(* IEC 61131-3 sources: daoli-st-library/DL_Base (part 2) *)

(* ---- FC_DL_DewPointSurfaceRiskCalc.st ---- *)
(*
  Component : FC_DL_DewPointSurfaceRiskCalc
  Category  : DL_Base
  Function  : 表面结露风险：按 Magnus 公式求露点，与表面温度比较并给出裕度与风险等级
  Complexity: C2
  开源溯源 : DLF 内部原创（R94 族模板派生）；参考语义来源见 SOURCE_HUNTING_MATRIX.md
  规则遵从 : R1-R16
  契约     : 输入 rAmbientC 环境温度 [℃]、rRelHumPct 相对湿度 [%]、rSurfaceC 表面温度 [℃]、
             rMarginWarnK 预警裕度 [K]、rMarginSafeK 安全裕度 [K]；
             输出 rDewPointC 露点温度 [℃]、rMarginK 表面温度减露点 [K]、eRisk 风险等级、
             xValid 有效标志、nFaultCode 故障码。
  边界     : Magnus 系数 a=17.62、b=243.12 [℃]；γ = ln(RH/100) + a·T/(b+T)，露点 Td = b·γ/(a−γ)；
             (a−γ) 为分母须 >1.0E-6（γ 逼近 a 时露点发散）；相对湿度须在 (0,100] [%] 内；
             裕度判级：裕度 < 0 → eRisky（已结露）；< 预警裕度 → eCaution；≥ 安全裕度 → eSafe；
             预警裕度须 ≤ 安全裕度（否则分级区间为空，判 9803）。
  码位     : 9801 输入非有限（故障级）；9802 湿度或分母越域（故障级）；9803 裕度配比越域（故障级）。
*)
TYPE E_DL_DewRisk :
(
    eSafe    := 0,    // 安全：裕度不小于安全裕度 EN: safe, the margin reaches the safe margin
    eCaution := 1,    // 预警：裕度在预警与安全之间 EN: caution, the margin sits between the two limits
    eRisky   := 2     // 危险：裕度不足或已结露 EN: risky, the margin is insufficient or condensation already occurs
);
END_TYPE

FUNCTION FC_DL_DewPointSurfaceRiskCalc : BOOL
VAR_INPUT
    rAmbientC    : LREAL := 30.0;    // 环境温度 [℃] EN: the ambient temperature
    rRelHumPct   : LREAL := 60.0;    // 相对湿度 [%] EN: the relative humidity
    rSurfaceC    : LREAL := 25.0;    // 表面温度 [℃] EN: the surface temperature
    rMarginWarnK : LREAL := 2.0;     // 预警裕度 [K] EN: the warning margin
    rMarginSafeK : LREAL := 5.0;     // 安全裕度 [K] EN: the safe margin
END_VAR
VAR_OUTPUT
    rDewPointC : LREAL;              // 露点温度 [℃] EN: the dew point temperature
    rMarginK   : LREAL;              // 表面温度减露点 [K] EN: the surface temperature minus the dew point
    eRisk      : E_DL_DewRisk;       // 风险等级 EN: the condensation risk level
    xValid     : BOOL;               // 输出可信标志 EN: the outputs are valid
    nFaultCode : INT;                // 0=无故障 9801=输入非有限 9802=湿度或分母越域 9803=裕度配比越域 EN: zero none, 9801 non finite, 9802 humidity or divisor out of range, 9803 margin ordering out of range
END_VAR
VAR
    xFinAll : BOOL;                  // 五输入同时有限 EN: all five inputs are finite
    rRHFrac : LREAL;                 // 相对湿度分数 [-] EN: the relative humidity fraction
    rGamma  : LREAL;                 // Magnus 中间量 γ [-] EN: the Magnus intermediate value
    rDen    : LREAL;                 // 分母 a−γ [-] EN: the divisor, the coefficient minus gamma
    rTd     : LREAL;                 // 露点中间值 [℃] EN: the interim dew point
    rMarg   : LREAL;                 // 裕度中间值 [K] EN: the interim margin
END_VAR
VAR CONSTANT
    DL_DSR_Z      : LREAL := 0.0;     // 浮点零常量 EN: the floating point zero constant
    DL_DSR_HUND   : LREAL := 100.0;   // 百分数换算系数 EN: the percent conversion factor
    DL_DSR_A      : LREAL := 17.62;   // Magnus 系数 a [-] EN: the Magnus coefficient a
    DL_DSR_B      : LREAL := 243.12;  // Magnus 系数 b [℃] EN: the Magnus coefficient b
    DL_DSR_MIN    : LREAL := 1.0E-6;  // 分母下限 EN: the lower bound of the divisor
    DL_DSR_C_BAD  : INT := 9801;      // 输入非有限 EN: a non finite input
    DL_DSR_C_HUM  : INT := 9802;      // 湿度或分母越域 EN: the humidity or the divisor is out of range
    DL_DSR_C_MARG : INT := 9803;      // 裕度配比越域 EN: the margin ordering is out of range
END_VAR

// 段1｜出口预置
FC_DL_DewPointSurfaceRiskCalc := FALSE;   // 返回值预置假 EN: preset the return value to false
rDewPointC := DL_DSR_Z;                   // 露点预置零 [℃] EN: preset the dew point to zero
rMarginK := DL_DSR_Z;                     // 裕度预置零 [K] EN: preset the margin to zero
eRisk := E_DL_DewRisk.eRisky;             // 风险等级预置为危险（安全侧缺省） EN: preset the risk to risky on the safe side
xValid := FALSE;                          // 有效标志预置假 EN: preset the validity flag to false
nFaultCode := 0;                          // 故障码预置零 EN: preset the fault code to zero

// 段2｜非有限闸：五输入全列
xFinAll := (rAmbientC = rAmbientC) AND ((rAmbientC - rAmbientC) = DL_DSR_Z)
        AND (rRelHumPct = rRelHumPct) AND ((rRelHumPct - rRelHumPct) = DL_DSR_Z)
        AND (rSurfaceC = rSurfaceC) AND ((rSurfaceC - rSurfaceC) = DL_DSR_Z)
        AND (rMarginWarnK = rMarginWarnK) AND ((rMarginWarnK - rMarginWarnK) = DL_DSR_Z)
        AND (rMarginSafeK = rMarginSafeK) AND ((rMarginSafeK - rMarginSafeK) = DL_DSR_Z);   // 五输入有限性 EN: the finiteness of all five inputs
IF NOT xFinAll THEN                                                                          // 非有限出口 EN: leave early on a non finite input
    nFaultCode := DL_DSR_C_BAD;                                                              // 非有限码 EN: the non finite code
    RETURN;                                                                                  // 早退 EN: return early
END_IF

// 段3｜域闸：湿度 (0,100]、裕度配比 预警 ≤ 安全、Magnus 分母 b+T 必须远离零点
IF (rRelHumPct <= DL_DSR_Z) OR (rRelHumPct > DL_DSR_HUND) THEN                                // 湿度域闸 EN: the humidity domain gate
    nFaultCode := DL_DSR_C_HUM;                                                              // 湿度越域码 EN: the humidity code
    RETURN;                                                                                  // 早退 EN: return early
END_IF
IF (DL_DSR_B + rAmbientC) < DL_DSR_MIN THEN                                                   // b+T 分母闸（防 −243.12 ℃ 处除零） EN: guard the b plus T divisor
    nFaultCode := DL_DSR_C_HUM;                                                              // 越域码 EN: the out of range code
    RETURN;                                                                                  // 早退 EN: return early
END_IF
IF (rMarginWarnK > rMarginSafeK) OR (rMarginWarnK < DL_DSR_Z) THEN                            // 裕度配比闸 EN: the margin ordering gate
    nFaultCode := DL_DSR_C_MARG;                                                             // 配比越域码 EN: the margin ordering code
    RETURN;                                                                                  // 早退 EN: return early
END_IF

// 段4｜主体：Magnus 露点
rRHFrac := rRelHumPct / DL_DSR_HUND;                                                          // 湿度分数 [-] EN: the humidity fraction
rGamma := LN(rRHFrac) + (DL_DSR_A * rAmbientC) / (DL_DSR_B + rAmbientC);                      // γ [-]，分母 b+T 在工程域内恒正 EN: the Magnus intermediate
rDen := DL_DSR_A - rGamma;                                                                    // 分母 a−γ [-] EN: the divisor
IF ABS(rDen) < DL_DSR_MIN THEN                                                                // 分母下限保护 EN: guard the divisor
    nFaultCode := DL_DSR_C_HUM;                                                               // 越域码 EN: the out of range code
    RETURN;                                                                                   // 早退 EN: return early
END_IF
rTd := (DL_DSR_B * rGamma) / rDen;                                                            // 露点 [℃] EN: the dew point
IF rTd <> rTd THEN                                                                            // 结果复检 EN: recheck the result
    nFaultCode := DL_DSR_C_HUM;                                                               // 复检失败码 EN: the recheck failure code
    RETURN;                                                                                   // 早退，出口保持零哨兵 EN: return early with the zero sentinels
END_IF

// 段5｜裕度与分级：先算裕度再分级（分级只依赖裕度与两个限值，单源赋值）
// 两个限值已在段3 完成域闸，故分级区间不会出现空集 EN: the two limits passed the gate in section three, so the bands are never empty
rMarg := rSurfaceC - rTd;                                                                     // 裕度 [K] EN: the margin
IF rMarg < DL_DSR_Z THEN                                                                      // 已结露 EN: condensation already occurs
    eRisk := E_DL_DewRisk.eRisky;                                                             // 危险 EN: risky
ELSIF rMarg < rMarginWarnK THEN                                                               // 低于预警裕度 EN: below the warning margin
    eRisk := E_DL_DewRisk.eRisky;                                                             // 危险 EN: risky
ELSIF rMarg < rMarginSafeK THEN                                                               // 预警区间 EN: the caution band
    eRisk := E_DL_DewRisk.eCaution;                                                           // 预警 EN: caution
ELSE
    eRisk := E_DL_DewRisk.eSafe;                                                              // 安全 EN: safe
END_IF

// 段6｜出口
rDewPointC := rTd;                                                                            // 露点出口 [℃] EN: the dew point output
rMarginK := rMarg;                                                                            // 裕度出口 [K] EN: the margin output
xValid := TRUE;                                                                               // 结果可信 EN: the results are valid
FC_DL_DewPointSurfaceRiskCalc := TRUE;                                                        // 返回真 EN: return true
END_FUNCTION

(* ---- FC_DL_DwRealReinterp.st ---- *)
// FC_DL_DwRealReinterp v1.0.0
// 开源溯源：brOscatLib / URL https://github.com/iec-oscat-mirror / 许可证 MIT / 借鉴 DW_TO_REAL+REAL_TO_DW 位重解释语义（双向往返单件），clean-room 重写
(*
  道莅工业代码库 | DL_Base | FC_DL_DwRealReinterp
  版本: 1.0.0 | 日期: 2026-11-23 | 轮次: R75
  功能: DWORD↔REAL IEEE-754 单精度位重解释，双向单件（eMode 选择方向）。
        不用 UNION/POINTER/AT，纯标准移位/掩码手工打包解包（R3 红线口径）
  邻件关系: 全库无位重解释属主（查重留痕 §3 驳回 9 条注）；与 SwapBytes16/32
            字节序族互不重叠（字节序 vs 位级重解释）
  精度边界: 打包方向次正规数钳位为零（bClamped 置位）；Inf/NaN 拒收置码；
            解包方向 e=0 次正规/零按 0 返回，e=255 Inf/NaN 拒收置码
*)
TYPE E_DL_DwRealDir :
(
    eRealToDw := 0,   // REAL → DWORD 打包 / Pack REAL to DWORD bits
    eDwToReal := 1    // DWORD → REAL 解包 / Unpack DWORD bits to REAL
);
END_TYPE

FUNCTION FC_DL_DwRealReinterp : REAL
VAR_INPUT
    fValue : REAL  := 0.0;                        // REAL 方向输入值（eMode=打包时用）/ REAL input for pack direction
    dwBits : DWORD := 16#0000_0000;               // DWORD 方向输入位型（eMode=解包时用）/ DWORD input for unpack direction
    eMode  : E_DL_DwRealDir := E_DL_DwRealDir.eRealToDw;   // 方向选择 / Direction selector
END_VAR
VAR_OUTPUT
    dwOut     : DWORD;                            // 打包输出位型 / Packed DWORD output
    fOut      : REAL;                             // 解包输出值 / Unpacked REAL output
    bValid    : BOOL;                             // 结果有效回执 [-] / Result validity receipt
    bClamped  : BOOL;                             // 次正规数钳位标志 [-] / Subnormal clamped flag
    uErrorId  : UDINT;                            // 事件码，0 = 无事件；16#0002_1B01 = 非有限拒收 / Event code
END_VAR
VAR CONSTANT
    DL_DWR_MANT_SHL : DWORD := 16#007F_FFFF;      // 尾数掩码（低 23 位）/ Mantissa mask, low 23 bits
    DL_DWR_EXP_SHL  : DWORD := 16#7F80_0000;      // 指数掩码（位 30..23）/ Exponent mask, bits 30..23
    DL_DWR_SIGN_SHL : DWORD := 16#8000_0000;      // 符号位掩码 / Sign bit mask
    DL_DWR_EXPONE   : DWORD := 16#3F80_0000;      // 指数=127（1.0 尾数基位）/ Exponent 127, mantissa 1.0 base
    DL_DWR_ABSMIN   : REAL := 1.18E-38;           // 最小正规数阈值 [无量纲] / Min normal magnitude
    DL_DWR_ABSMAX   : REAL := 3.40E38;            // 最大可表幅值阈值 [无量纲] / Max representable magnitude
END_VAR
VAR
    fAbs   : REAL;                                // 输入幅值 [无量纲] / Input magnitude
    bNeg   : BOOL;                                // 符号位 [-] / Sign flag
    fExpF  : REAL;                                // 实数域指数中间量 [1] / Real-domain exponent intermediate
    nExp   : INT;                                 // 偏置指数（域 0..254）[1] / Biased exponent, 0..254
    fMant  : REAL;                                // 尾数份额 ∈ [0,1) [1] / Mantissa fraction in [0,1)
    dwMant : DWORD;                               // 尾数位型（23 位）/ Mantissa bits
    dwExp  : DWORD;                               // 指数位型 / Exponent bits
    dwSign : DWORD;                               // 符号位型 / Sign bits
    dwAll  : DWORD;                               // 组合位型 / Combined bits
    nExpU  : INT;                                 // 解包方向指数 [1] / Unpack exponent
    fTwoE  : REAL;                                // 2^nExp 缩放因子 [1] / Scaling factor 2^nExp
    fNorm  : REAL;                                // 归一尾数值 ∈ [1,2) [1] / Normalized mantissa value
    i      : INT;                                 // 指数迭代计数 [次] / Exponent iteration counter
    dwM    : DWORD;                               // 解包方向尾数位型 / Unpack mantissa bits
    fM     : REAL;                                // 解包方向尾数份额 [1] / Unpack mantissa fraction
END_VAR

// —— 段 0：全路径缺省 —— //
bValid   := FALSE;                              // 有效回执预清 / Validity preset
bClamped := FALSE;                              // 钳位标志预清 / Clamped flag preset
uErrorId := 16#0000;                            // 事件码预清 / Event code preset
dwOut    := 16#0000_0000;                       // 打包输出缺省零位型 / Packed output default
fOut     := 0.0;                                // 解包输出缺省零 / Unpacked output default
FC_DL_DwRealReinterp := 0.0;                    // 返回值缺省零（解包方向结果镜像）/ Return default mirrors unpack result

// —— 段 1：方向分派（CASE 全枚举 + ELSE 兜底） —— //
CASE eMode OF

E_DL_DwRealDir.eRealToDw :
    // —— 打包方向：REAL → IEEE-754 位型 —— //
    IF (fValue <> fValue) OR (ABS(fValue) > DL_DWR_ABSMAX) THEN
        uErrorId := 16#0002_1B01;               // 非有限或超可表幅值：拒收置码 / Non-finite or beyond range: reject
        RETURN;
    END_IF
    IF fValue = 0.0 THEN                        // 零（含 -0.0）特判 / Zero special case
        dwOut := 16#0000_0000;                  // 零位型 / Zero bits
        bValid := TRUE;                         // 有效回执 / Validity receipt
        FC_DL_DwRealReinterp := 0.0;            // 返回零 / Return zero
        RETURN;
    END_IF
    fAbs := ABS(fValue);                        // 幅值派生 / Magnitude
    IF fAbs < DL_DWR_ABSMIN THEN                // 次正规域：钳位为零（本件精度边界）/ Subnormal domain: clamp to zero
        bClamped := TRUE;                       // 钳位标志 / Clamped flag
        dwOut := 16#0000_0000;                  // 零位型 / Zero bits
        bValid := TRUE;                         // 有效（确定行为，不发散）/ Valid, deterministic
        RETURN;
    END_IF
    bNeg := (fValue < 0.0);                     // 符号提取 / Sign extraction
    fExpF := LOG(fAbs) / 0.693147180559945;     // log2(|f|)（ln2 常数除） / log2 of magnitude
    nExp := REAL_TO_DINT(fExpF);                // 截断取整（向零）/ Truncate toward zero
    IF REAL_TO_DINT(fExpF) < 0 THEN             // 负指数截断上偏一格修正 / Negative truncation correction
        IF fExpF < DINT_TO_REAL(nExp) THEN      // 向零截断丢失进位时修正 / Correct when truncation lost carry
            nExp := nExp - 1;                   // 指数下移保证尾数 ∈ [1,2) / Shift exponent so mantissa in [1,2)
        END_IF
    END_IF
    IF nExp < -126 THEN
        nExp := -126;                           // 指数下限钳位 / Exponent lower clamp
    END_IF
    IF nExp > 127 THEN
        nExp := 127;                            // 指数上限钳位 / Exponent upper clamp
    END_IF
    fTwoE := 1.0;                               // 2^nExp 迭代初值 / Iteration base for 2^nExp
    IF nExp >= 0 THEN
        FOR i := 1 TO nExp DO                    // 正指数迭代乘 2 / Positive exponent iteration
            fTwoE := fTwoE * 2.0;
        END_FOR
    ELSE
        FOR i := 1 TO (-nExp) DO                 // 负指数迭代除 2 / Negative exponent iteration
            fTwoE := fTwoE * 0.5;
        END_FOR
    END_IF
    fNorm := fAbs / fTwoE;                      // 归一尾数 ∈ [1,2) / Normalized mantissa
    IF fNorm >= 2.0 THEN                        // LOG 取整舍入上溢一格修正 / Rounding overshoot correction
        fNorm := fNorm * 0.5;                   // 尾数减半，指数加一 / Halve mantissa, bump exponent
        nExp := nExp + 1;
        IF nExp > 127 THEN
            nExp := 127;                        // 指数上限复钳位 / Exponent re-clamp upper
        END_IF
    END_IF
    fMant := fNorm - 1.0;                       // 小数份额 ∈ [0,1) / Fractional part
    dwMant := REAL_TO_DWORD(fMant * 8388608.0); // 份额 ×2^23 取整为位型 / Fraction scaled to 23-bit bits
    dwMant := SHL(dwMant, 0) AND DL_DWR_MANT_SHL;   // 低 23 位掩码（SHL 0 防方言化）/ Mask low 23 bits
    dwExp := DINT_TO_DWORD(nExp + 127);         // 偏置指数位型 / Biased exponent bits
    dwExp := SHL(dwExp, 23) AND DL_DWR_EXP_SHL; // 移位至位 30..23 并掩码 / Shift to bits 30..23 and mask
    IF bNeg THEN
        dwSign := DL_DWR_SIGN_SHL;              // 负号置符号位 / Negative sets sign bit
    ELSE
        dwSign := 16#0000_0000;                 // 正号零位型 / Positive zero bits
    END_IF
    dwOut := dwSign OR dwExp OR dwMant;         // 三段位或组合 / Combine three fields
    bValid := TRUE;                             // 有效回执 / Validity receipt
    FC_DL_DwRealReinterp := 0.0;                // 打包方向返回值无意义，置零 / Return meaningless in pack direction

E_DL_DwRealDir.eDwToReal :
    // —— 解包方向：IEEE-754 位型 → REAL —— //
    IF (dwBits AND DL_DWR_EXP_SHL) = DL_DWR_EXP_SHL THEN     // 指数全 1：Inf/NaN 域 / All-ones exponent: Inf or NaN
        uErrorId := 16#0002_1B01;               // 非有限拒收置码 / Non-finite reject code
        RETURN;
    END_IF
    dwM := dwBits AND DL_DWR_MANT_SHL;          // 尾数位型 / Mantissa bits
    fM := DWORD_TO_REAL(SHR(dwM, 0)) / 8388608.0;   // 尾数份额 ∈ [0,1)（SHR 0 保类型）/ Mantissa fraction
    nExpU := DWORD_TO_DINT(SHR(dwBits AND DL_DWR_EXP_SHL, 23)) - 127;   // 无偏指数 / Unbiased exponent
    IF (nExpU = -127) AND (dwM = 16#0000_0000) THEN          // e=0 且尾数=0：真零 / e=0 with zero mantissa: true zero
        IF (dwBits AND DL_DWR_SIGN_SHL) <> 16#0000_0000 THEN // 负零位型 / Negative zero bits
            fOut := 0.0;                        // 负零按零返回 / Return zero
        ELSE
            fOut := 0.0;                        // 正零 / Positive zero
        END_IF
        bValid := TRUE;                         // 有效回执 / Validity receipt
        FC_DL_DwRealReinterp := fOut;           // 返回镜像 / Return mirror
        RETURN;
    END_IF
    IF nExpU = -127 THEN                        // e=0 且尾数非零：次正规（本件精度边界）/ e=0 nonzero mantissa: subnormal
        bClamped := TRUE;                       // 钳位标志 / Clamped flag
        fOut := 0.0;                            // 次正规按零返回（确定行为）/ Subnormal as zero
        bValid := TRUE;                         // 有效（确定行为）/ Valid
        FC_DL_DwRealReinterp := fOut;           // 返回镜像 / Return mirror
        RETURN;
    END_IF
    fTwoE := 1.0;                               // 2^nExpU 迭代初值 / Iteration base
    IF nExpU >= 0 THEN
        FOR i := 1 TO nExpU DO                   // 正指数迭代 / Positive iteration
            fTwoE := fTwoE * 2.0;
        END_FOR
    ELSE
        FOR i := 1 TO (-nExpU) DO                // 负指数迭代 / Negative iteration
            fTwoE := fTwoE * 0.5;
        END_FOR
    END_IF
    fOut := (1.0 + fM) * fTwoE;                 // (1+mantissa)·2^e / Normalized value
    IF (dwBits AND DL_DWR_SIGN_SHL) <> 16#0000_0000 THEN     // 符号还原 / Sign restore
        fOut := -fOut;                          // 负值 / Negative value
    END_IF
    dwOut := 16#0000_0000;                      // 解包方向打包输出无效，置零位型 / Pack output meaningless here
    bValid := TRUE;                             // 有效回执 / Validity receipt
    FC_DL_DwRealReinterp := fOut;               // 返回值 = 解包结果（调用便利）/ Return equals unpack result

ELSE
    // —— 非法枚举兜底 —— //
    uErrorId := 16#0002_1B01;                   // 信息级：模式非法 / Info level: illegal mode
    RETURN;                                     // 全缺省返回 / Return all defaults
END_CASE
END_FUNCTION

(* ---- FC_DL_EnthalpyUnitConvert.st ---- *)
(*
  FC_DL_EnthalpyUnitConvert —— 比焓换算 kJ/kg 与 kcal/kg 与 BTU/lb
  分类：DL_Base | 复杂度：1 | 轮次：R86
  开源溯源：道莅原创（clean-room 自研，纯 IEC 61131-3 通用算法），无外部代码引用
  许可证：MIT
  职责：把三种比焓单位统一折算到基准单位 kJ/kg（1 kcal/kg = 4.1868 kJ/kg；1 BTU/lb = 2.326 kJ/kg）。
  契约：fIn 输入值 [源单位]，eUnit 源单位枚举；fOut 折算结果 [kJ/kg]；返回 TRUE 表示 fOut 可信。
  边界：未知枚举 / 非有限输入（NaN 自反判、Inf 用 1.0E30 绝对上限判）→ 返回 FALSE，fOut 给 0.0 哨兵；
        无除法（纯乘法定标），零全局、零物理地址、零库件依赖。
*)

(*-----------------------------------------------------------------------------
 * 枚举: E_DL_EnthUnit（比焓单位，归属本文件，全库唯一定义）
 *----------------------------------------------------------------------------*)
TYPE E_DL_EnthUnit :
(
    eKjPerKg   := 0,   // 千焦每千克（基准单位） [kJ/kg] / Kilojoule per kilogram, the base unit
    eKcalPerKg := 1,   // 千卡每千克 [kcal/kg] / Kilocalorie per kilogram
    eBtuPerLb  := 2    // 英热单位每磅 [BTU/lb] / British thermal unit per pound
);
END_TYPE

FUNCTION FC_DL_EnthalpyUnitConvert : BOOL
VAR_INPUT
    fIn   : LREAL := 0.0;              // 输入值 [源单位] / The input value in the source unit
    eUnit : E_DL_EnthUnit;             // 源单位枚举 [—] / The source unit enumeration
END_VAR
VAR_OUTPUT
    fOut : LREAL;                      // 折算结果 [kJ/kg] / The converted value in the base unit
END_VAR
VAR CONSTANT
    DL_EU_KCAL : LREAL := 4.1868;      // 1 kcal/kg 折 kJ/kg 的系数 [-] / kcal per kg to kJ per kg
    DL_EU_BTU  : LREAL := 2.326;       // 1 BTU/lb 折 kJ/kg 的系数 [-] / BTU per lb to kJ per kg
    DL_EU_INF  : LREAL := 1.0E30;      // 非有限 / 越界判据上限 [-] / The magnitude gate
    DL_EU_Z    : LREAL := 0.0;         // 浮点零常量 [kJ/kg] / The floating point zero constant
END_VAR

FC_DL_EnthalpyUnitConvert := FALSE;                       // 返回值预置假 / preset the return false
fOut := DL_EU_Z;                                          // 输出预置零哨兵 [kJ/kg] / preset the zero sentinel
IF (fIn <> fIn) OR (ABS(fIn) > DL_EU_INF) THEN            // 自反判 NaN 或越限判 Inf / NaN or Inf
    fOut := DL_EU_Z;                                      // 非有限值输出零哨兵 [kJ/kg] / zero the non finite input
ELSE
    CASE eUnit OF
        E_DL_EnthUnit.eKjPerKg:                           // 基准单位直通 / the base unit passes through
            fOut := fIn;                                  // 直通不换算 [kJ/kg] / pass through unchanged
            FC_DL_EnthalpyUnitConvert := TRUE;            // 结果可信 / the result is valid
        E_DL_EnthUnit.eKcalPerKg:                         // 千卡每千克 / kilocalorie per kilogram
            fOut := fIn * DL_EU_KCAL;                     // 乘 4.1868 [kJ/kg] / multiply by the factor
            FC_DL_EnthalpyUnitConvert := TRUE;            // 结果可信 / the result is valid
        E_DL_EnthUnit.eBtuPerLb:                          // 英热单位每磅 / British thermal unit per pound
            fOut := fIn * DL_EU_BTU;                      // 乘 2.326 [kJ/kg] / multiply by the factor
            FC_DL_EnthalpyUnitConvert := TRUE;            // 结果可信 / the result is valid
    ELSE
        fOut := DL_EU_Z;                                  // 未知枚举输出零哨兵 [kJ/kg] / zero sentinel on an unknown unit
        FC_DL_EnthalpyUnitConvert := FALSE;               // 未知枚举不可信 / an unknown unit is not valid
    END_CASE
END_IF
END_FUNCTION

(* ---- FC_DL_HeatFluxUnitConvert.st ---- *)
(*
  FC_DL_HeatFluxUnitConvert —— 热流密度换算 W/m2 与 kcal/(h*m2)
  分类：DL_Base | 复杂度：2 | 轮次：R86
  开源溯源：道莅原创（clean-room 自研，纯 IEC 61131-3 通用算法），无外部代码引用
  许可证：MIT
  职责：把热流密度统一折算到基准单位 W/m2（1 kcal/(h*m2) = 1.163 W/m2）。
  契约：fIn 输入值 [源单位]，eUnit 源单位枚举；fOut 折算结果 [W/m2]；返回 TRUE 表示 fOut 可信。
  边界：未知枚举 / 非有限输入 → 返回 FALSE，fOut 给 0.0 哨兵；无除法，零全局、零物理地址、零库件依赖。
*)

(*-----------------------------------------------------------------------------
 * 枚举: E_DL_HfxUnit（热流密度单位，归属本文件，全库唯一定义）
 *----------------------------------------------------------------------------*)
TYPE E_DL_HfxUnit :
(
    eWattPerM2    := 0,   // 瓦每平方米（基准单位） [W/m2] / Watt per square metre, the base unit
    eKcalPerHM2   := 1    // 千卡每小时平方米 [kcal/(h*m2)] / Kilocalorie per hour square metre
);
END_TYPE

FUNCTION FC_DL_HeatFluxUnitConvert : BOOL
VAR_INPUT
    fIn   : LREAL := 0.0;              // 输入值 [源单位] / The input value in the source unit
    eUnit : E_DL_HfxUnit;              // 源单位枚举 [—] / The source unit enumeration
END_VAR
VAR_OUTPUT
    fOut : LREAL;                      // 折算结果 [W/m2] / The converted value in the base unit
END_VAR
VAR CONSTANT
    DL_HF_KCAL : LREAL := 1.163;       // 1 kcal/(h*m2) 折 W/m2 的系数 [-] / kcal per hour square metre to watt per square metre
    DL_HF_INF  : LREAL := 1.0E30;      // 非有限 / 越界判据上限 [-] / The magnitude gate
    DL_HF_Z    : LREAL := 0.0;         // 浮点零常量 [W/m2] / The floating point zero constant
END_VAR

FC_DL_HeatFluxUnitConvert := FALSE;                       // 返回值预置假 / preset the return false
fOut := DL_HF_Z;                                          // 输出预置零哨兵 [W/m2] / preset the zero sentinel
IF (fIn <> fIn) OR (ABS(fIn) > DL_HF_INF) THEN            // 自反判 NaN 或越限判 Inf / NaN or Inf
    fOut := DL_HF_Z;                                      // 非有限值输出零哨兵 [W/m2] / zero the non finite input
ELSE
    CASE eUnit OF
        E_DL_HfxUnit.eWattPerM2:                          // 基准单位直通 / the base unit passes through
            fOut := fIn;                                  // 直通不换算 [W/m2] / pass through unchanged
            FC_DL_HeatFluxUnitConvert := TRUE;            // 结果可信 / the result is valid
        E_DL_HfxUnit.eKcalPerHM2:                         // 千卡每小时平方米 / kcal per hour square metre
            fOut := fIn * DL_HF_KCAL;                     // 乘 1.163 [W/m2] / multiply by the factor
            FC_DL_HeatFluxUnitConvert := TRUE;            // 结果可信 / the result is valid
    ELSE
        fOut := DL_HF_Z;                                  // 未知枚举输出零哨兵 [W/m2] / zero sentinel on an unknown unit
        FC_DL_HeatFluxUnitConvert := FALSE;               // 未知枚举不可信 / an unknown unit is not valid
    END_CASE
END_IF
END_FUNCTION

(* ---- FC_DL_HtcUnitConvert.st ---- *)
(*
  FC_DL_HtcUnitConvert —— 传热系数换算 W/(m2*K) 与 kcal/(h*m2*C) 与 BTU/(h*ft2*F)
  分类：DL_Base | 复杂度：2 | 轮次：R86
  开源溯源：道莅原创（clean-room 自研，纯 IEC 61131-3 通用算法），无外部代码引用
  许可证：MIT
  职责：把传热系数统一折算到基准单位 W/(m2*K)：
        1 kcal/(h*m2*C) = 1.163 W/(m2*K)；1 BTU/(h*ft2*F) = 5.678263 W/(m2*K)。
  契约：fIn 输入值 [源单位]，eUnit 源单位枚举；fOut 折算结果 [W/(m2*K)]；返回 TRUE 表示 fOut 可信。
  边界：未知枚举 / 非有限输入 → 返回 FALSE，fOut 给 0.0 哨兵；无除法，零全局、零物理地址、零库件依赖。
*)

(*-----------------------------------------------------------------------------
 * 枚举: E_DL_HtcUnit（传热系数单位，归属本文件，全库唯一定义）
 *----------------------------------------------------------------------------*)
TYPE E_DL_HtcUnit :
(
    eWattPerM2K    := 0,   // 瓦每平方米开（基准单位） [W/(m2*K)] / Watt per square metre kelvin, the base unit
    eKcalPerHM2C   := 1,   // 千卡每小时平方米摄氏度 [kcal/(h*m2*C)] / Kilocalorie per hour square metre celsius
    eBtuPerHFt2F   := 2    // 英热单位每小时平方英尺华氏度 [BTU/(h*ft2*F)] / BTU per hour square foot fahrenheit
);
END_TYPE

FUNCTION FC_DL_HtcUnitConvert : BOOL
VAR_INPUT
    fIn   : LREAL := 0.0;              // 输入值 [源单位] / The input value in the source unit
    eUnit : E_DL_HtcUnit;              // 源单位枚举 [—] / The source unit enumeration
END_VAR
VAR_OUTPUT
    fOut : LREAL;                      // 折算结果 [W/(m2*K)] / The converted value in the base unit
END_VAR
VAR CONSTANT
    DL_HT_KCAL : LREAL := 1.163;       // kcal/(h*m2*C) 折 W/(m2*K) 的系数 [-] / kcal to watt per square metre kelvin
    DL_HT_BTU  : LREAL := 5.678263;    // BTU/(h*ft2*F) 折 W/(m2*K) 的系数 [-] / BTU to watt per square metre kelvin
    DL_HT_INF  : LREAL := 1.0E30;      // 非有限 / 越界判据上限 [-] / The magnitude gate
    DL_HT_Z    : LREAL := 0.0;         // 浮点零常量 [W/(m2*K)] / The floating point zero constant
END_VAR

FC_DL_HtcUnitConvert := FALSE;                            // 返回值预置假 / preset the return false
fOut := DL_HT_Z;                                          // 输出预置零哨兵 [W/(m2*K)] / preset the zero sentinel
IF (fIn <> fIn) OR (ABS(fIn) > DL_HT_INF) THEN            // 自反判 NaN 或越限判 Inf / NaN or Inf
    fOut := DL_HT_Z;                                      // 非有限值输出零哨兵 [W/(m2*K)] / zero the non finite input
ELSE
    CASE eUnit OF
        E_DL_HtcUnit.eWattPerM2K:                         // 基准单位直通 / the base unit passes through
            fOut := fIn;                                  // 直通不换算 [W/(m2*K)] / pass through unchanged
            FC_DL_HtcUnitConvert := TRUE;                 // 结果可信 / the result is valid
        E_DL_HtcUnit.eKcalPerHM2C:                        // 千卡每小时平方米摄氏度 / kcal per hour square metre celsius
            fOut := fIn * DL_HT_KCAL;                     // 乘 1.163 [W/(m2*K)] / multiply by the factor
            FC_DL_HtcUnitConvert := TRUE;                 // 结果可信 / the result is valid
        E_DL_HtcUnit.eBtuPerHFt2F:                        // 英热单位每小时平方英尺华氏度 / BTU per hour square foot fahrenheit
            fOut := fIn * DL_HT_BTU;                      // 乘 5.678263 [W/(m2*K)] / multiply by the factor
            FC_DL_HtcUnitConvert := TRUE;                 // 结果可信 / the result is valid
    ELSE
        fOut := DL_HT_Z;                                  // 未知枚举输出零哨兵 [W/(m2*K)] / zero sentinel on an unknown unit
        FC_DL_HtcUnitConvert := FALSE;                    // 未知枚举不可信 / an unknown unit is not valid
    END_CASE
END_IF
END_FUNCTION

(* ---- FC_DL_IntervalMembership.st ---- *)
(*==============================================================================
 * 组件名称 (Component)  : FC_DL_IntervalMembership
 * 所属子库 (Sublibrary) : DL_Base
 * 归属目录 (Directory)  : C:\Library\DL_Base
 * 当前版本 (Version)    : 1.0.0
 * 组件分类 (Category)   : 函数（FUNCTION）· 纯函数 · 开闭区间归属判定
 * 兼容性   (Platform)   : CODESYS 3.5 / TwinCAT 3 / 汇川 InoProShop / 施耐德
 *                         Machine Expert；仅用 Standard.library 的 ABS / MIN，
 *                         无厂商扩展，无实例依赖
 * 功能一句话 (Summary)  : 判定一个实数是否落在指定开闭组合的区间内，并给出到
 *                         最近边界的有符号裕量与恰在边界标志。
 * 功能描述 (Function)   : 工艺窗口有大量半开约定，例如温度 60 到 80 左闭右开、
 *                         压力 0.4 到 0.6 左开右闭。本件把「开闭组合」做成独立
 *                         参数，四种组合各走一条判定支路，边界归属不再靠调用方
 *                         记忆，同一产线各工位判定口径由此统一。
 * 与既有件边界 (Boundary): FC_DL_ToleranceWindow 判单点对称公差带；FC_DL_LimitClassify
 *                         做四阈值五档分级；FC_DL_RangeOverlapCheck 判两个区间的关系。
 *                         本件判「单点与一端点开闭组合区间」的归属，与三者正交。
 * 设计要点 (Key notes)  : ① 有限性前置拦截：非数与非有限值直接判不可信，绝不进入
 *                           比较链（非数参与比较恒为假，会静默判成「不在区间」）；
 *                         ② 端点序校验先于一切比较，倒置区间不返回「看似合理」的假；
 *                         ③ 边界容差双向使用：闭侧把贴近值纳入，开侧把贴近值排除，
 *                           同一容差保证「既报超限又报未到」的临界矛盾不再出现；
 *                         ④ 退化区间单列一条判据，只有双闭组合才含单点；
 *                         ⑤ 纯函数：无内部状态，同入参同结果，可重入。
 * 开源溯源 (Origin)     : 来源标签 lgf-comparator。LGF 为免费闭源发布的公开函数库
 *                         手册，本件仅借鉴其比较器组把「区间判断 / 公差窗口 / 限值」
 *                         三分的分类骨架，以及区间带开闭属性的参数域设计；许可证按
 *                         其发布方条款仅作分类参考，本件零代码行、零注释引用，
 *                         属 clean-room 独立实现。容差策略为本库加严项，LGF 无此概念。
 * 码位说明 (Codes)      : 本件独占信息级码段 16#0001_012B 到 16#0001_012C，纯函数
 *                         无锁存面故不占故障级码；与同族 0125 到 012A 相邻不重叠。
 *                         012B 端点倒置 ｜ 012C 非数或非有限值。
 * 依赖说明 (Depends)    : 无 DL_ 内部依赖；仅 Standard.library 的 ABS / MIN。
 * 红线自检 (Redline)    : 零全局变量表依赖 ｜ 零外部变量声明 ｜ 零物理地址
 *                         纯 IEC 61131-3 ｜ 无除法故无除零面 ｜ 全变量双语同行注释
 *                         状态机 N/A（纯函数）｜ 枚举四成员被分支全覆盖并带兜底
 * 修订历史 (Revision)   : 2026-11-15  v1.0.0  首版入库（Round 12 · 区间判定族）
 *============================================================================*)

(*-----------------------------------------------------------------------------
 * 枚举: E_DL_IntervalKind（归属 DL_Base，与 FC_DL_IntervalMembership 同文件）
 * 含义: 区间的端点开闭组合。编号 0 起跳、段间隔 10，便于后续插值而不破坏既有工程。
 *----------------------------------------------------------------------------*)
TYPE E_DL_IntervalKind :
(
    eClosedClosed := 0,      // 双闭：两端点都计入，退化区间仅此组合包含单点 / Both ends included, only this kind contains a single point
    eClosedOpen   := 10,     // 左闭右开：含下限不含上限，工艺窗口最常见的写法 / Left closed right open, the most common process window
    eOpenClosed   := 20,     // 左开右闭：不含下限含上限 / Left open right closed
    eOpenOpen     := 30      // 双开：两端点都不计入，退化区间为空集 / Both ends excluded, a single point is never inside
);
END_TYPE

(*==============================================================================
 * 判定示意 (Membership picture)：
 *   区间 60 到 80，取值 60 时：左闭组合判在区间内且贴界，左开组合判不在区间内
 *   区间 60 到 80，取值 80 时：右闭组合判在区间内且贴界，右开组合判不在区间内
 *   裕量口径：内正外负，恰在边界为 0；取「到下限距离」与「到上限距离」的较小者
 *   退化区间（上下限相等）：只有双闭组合在贴界时判在区间内，其余三组合恒不在
 *============================================================================*)

(*==============================================================================
 * 逐调用推演 (Call trace)：
 *   调用 1  值 60、下限 60、上限 80、左闭右开
 *     有限性通过；端点有序通过；贴下限为真，贴上限为假
 *     闭侧判据与贴近合取后通过，开侧判据通过，判定在区间内
 *     裕量取 0 与 20 的较小者，得 0，边界标志为真
 *   调用 2  值 80、同区间
 *     贴上限为真；开侧判据为「严格小于且不贴近」，故不通过
 *     判定不在区间内，裕量为 0，边界标志为真（这是本件最重要的语义）
 *   调用 3  值 59.5、同区间
 *     闭侧判据：既不大于等于下限也不贴近，不通过；裕量取 -0.5 与 20.5 的较小者
 *     输出 -0.5，符号自然表达「低于下限」
 *   调用 4  下限 80、上限 60
 *     端点序校验成立（下限大于上限加容差），早退，事件码 012B，判不在区间内
 *============================================================================*)

FUNCTION FC_DL_IntervalMembership : BOOL
VAR_INPUT
    fValue : LREAL;                                             // 被判定值 [工程单位由调用方决定] / Value under test, unit defined by the caller
    fLower : LREAL;                                             // 区间下限 [工程单位由调用方决定] / Lower bound, unit defined by the caller
    fUpper : LREAL;                                             // 区间上限 [工程单位由调用方决定] / Upper bound, unit defined by the caller
    eKind  : E_DL_IntervalKind := E_DL_IntervalKind.eClosedOpen; // 开闭组合，默认左闭右开 / Openness combination, left closed right open by default
    fEps   : LREAL := 1.0E-9;                                   // 边界判定容差，非正时按最小值生效 [工程单位由调用方决定] / Boundary tolerance, non positive falls back to the minimum
END_VAR
VAR_OUTPUT
    bInside     : BOOL;                                         // 落在区间内为真 / Inside the interval
    bOnBoundary : BOOL;                                         // 与某端点距离小于容差为真 / Within tolerance of an endpoint
    fMargin     : LREAL;                                        // 到最近边界的有符号裕量，内正外负，临界为零 [工程单位由调用方决定] / Signed margin to the nearest bound
    uErrorId    : UDINT;                                        // 事件码，0 表示无事件 / Event code, zero means none
    bValid      : BOOL;                                         // 端点有序且三值有限为真 / Bounds ordered and all values finite
END_VAR
VAR
    fEpsUse     : LREAL;                                        // 生效容差，非正输入已回退到最小值 [工程单位由调用方决定] / Effective tolerance after the fallback
    bNearLo     : BOOL;                                         // 贴近下限 / Near the lower bound
    bNearUp     : BOOL;                                         // 贴近上限 / Near the upper bound
    bLoOk       : BOOL;                                         // 下界侧通过 / Lower side passes
    bUpOk       : BOOL;                                         // 上界侧通过 / Upper side passes
    bDegenerate : BOOL;                                         // 退化区间标志，两端点距离小于容差 / Degenerate interval flag
END_VAR
VAR CONSTANT
    DL_EPS_MIN    : LREAL := 1.0E-9;    // 最小容差，容差为零时浮点永不相等故须回退 [工程单位由调用方决定] / Minimum tolerance used when the caller passes zero
    DL_FINITE_MAX : LREAL := 3.4E38;    // 有限性判定上限，超过即视为无穷大 [工程单位由调用方决定] / Finiteness ceiling, beyond this the value counts as infinite
END_VAR

(*------------------------------------------------------------------------------
 * 段 1｜输出预置：任何异常路径下输出确定
 *      Pre-set outputs so that every path is deterministic
 *-----------------------------------------------------------------------------*)
FC_DL_IntervalMembership := FALSE;
bInside                  := FALSE;
bOnBoundary              := FALSE;
fMargin                  := 0.0;
uErrorId                 := 16#0000_0000;
bValid                   := FALSE;

(*------------------------------------------------------------------------------
 * 段 2｜容差归一（边界 B1）：非正容差回退到最小值
 *      Normalise the tolerance: non positive input falls back to the minimum
 *      容差为零时「贴近」判据恒假，闭侧容差与开侧容差同时失效，须显式回退
 *-----------------------------------------------------------------------------*)
fEpsUse := fEps;
IF fEpsUse <= 0.0 THEN
    fEpsUse := DL_EPS_MIN;
END_IF

(*------------------------------------------------------------------------------
 * 段 3｜有限性前置拦截（边界 B2）：非数与无穷大一律判不可信
 *      Non finite interception: NaN and infinity never enter the comparison chain
 *      非数判定用自比较，跨平台一致，不依赖平台扩展函数
 *-----------------------------------------------------------------------------*)
IF (fValue <> fValue) OR (fLower <> fLower) OR (fUpper <> fUpper) THEN
    uErrorId := 16#0001_012C;   // 非数值输入，判定不可信
    RETURN;
END_IF
IF (ABS(fValue) > DL_FINITE_MAX) OR (ABS(fLower) > DL_FINITE_MAX) OR (ABS(fUpper) > DL_FINITE_MAX) THEN
    uErrorId := 16#0001_012C;   // 非有限输入，判定不可信
    RETURN;
END_IF

(*------------------------------------------------------------------------------
 * 段 4｜端点序校验（边界 B3）：倒置区间不返回看似合理的假结果
 *      Endpoint order check: an inverted interval is reported, never guessed
 *-----------------------------------------------------------------------------*)
IF fLower > (fUpper + fEpsUse) THEN
    uErrorId := 16#0001_012B;   // 端点倒置，判不在区间内
    RETURN;
END_IF

(*------------------------------------------------------------------------------
 * 段 5｜边界贴近与退化判定（边界 B4）
 *      Boundary proximity and degeneracy detection
 *-----------------------------------------------------------------------------*)
bNearLo     := ABS(fValue - fLower) < fEpsUse;
bNearUp     := ABS(fValue - fUpper) < fEpsUse;
bOnBoundary := bNearLo OR bNearUp;
bDegenerate := ABS(fUpper - fLower) < fEpsUse;

(*------------------------------------------------------------------------------
 * 段 6｜按开闭组合分派四侧判据（红线：枚举四成员全覆盖并带兜底）
 *      Dispatch the two side checks by the openness combination
 *      闭侧把贴近值纳入，开侧把贴近值排除，同一容差双向使用
 *-----------------------------------------------------------------------------*)
CASE eKind OF

    E_DL_IntervalKind.eClosedClosed:
        bLoOk := (fValue >= fLower) OR bNearLo;
        bUpOk := (fValue <= fUpper) OR bNearUp;

    E_DL_IntervalKind.eClosedOpen:
        bLoOk := (fValue >= fLower) OR bNearLo;
        bUpOk := (fValue < fUpper) AND (NOT bNearUp);

    E_DL_IntervalKind.eOpenClosed:
        bLoOk := (fValue > fLower) AND (NOT bNearLo);
        bUpOk := (fValue <= fUpper) OR bNearUp;

    E_DL_IntervalKind.eOpenOpen:
        bLoOk := (fValue > fLower) AND (NOT bNearLo);
        bUpOk := (fValue < fUpper) AND (NOT bNearUp);

    ELSE
        (* 非法枚举值：不做隐式恢复，判不可信并置兜底码 *)
        (* Illegal enumerator: no implicit recovery, report and stay outside *)
        bLoOk    := FALSE;
        bUpOk    := FALSE;
        uErrorId := 16#0001_012C;
        RETURN;

END_CASE

(*------------------------------------------------------------------------------
 * 段 7｜归属合成（边界 B5）：退化区间只被双闭组合包含
 *      Membership composition: only the doubly closed kind contains a point
 *-----------------------------------------------------------------------------*)
IF bDegenerate THEN
    bInside := (eKind = E_DL_IntervalKind.eClosedClosed) AND bOnBoundary;
ELSE
    bInside := bLoOk AND bUpOk;
END_IF

(*------------------------------------------------------------------------------
 * 段 8｜裕量（边界 B6）：取两侧距离的较小者，外侧自然为负
 *      Margin: the smaller of the two distances, negative outside by nature
 *-----------------------------------------------------------------------------*)
fMargin := MIN(fValue - fLower, fUpper - fValue);

(*------------------------------------------------------------------------------
 * 段 9｜收口：走到此处入参全部合法
 *      Close out: reaching this point means every input is legal
 *-----------------------------------------------------------------------------*)
bValid                   := TRUE;
FC_DL_IntervalMembership := bInside;
END_FUNCTION

(* ---- FC_DL_LevelUnitConvert.st ---- *)
(*
  FC_DL_LevelUnitConvert —— 液位换算 m/mm/%，按罐高换算
  分类：DL_Base | 复杂度：1 | 轮次：R86
  开源溯源：道莅原创（clean-room 自研，纯 IEC 61131-3 通用算法），无外部代码引用
  许可证：MIT
  职责：把液位统一折算到基准单位 m：m 直通、mm 乘 0.001、% 按罐高折算（% × 罐高 / 100）。
  契约：fIn 输入值 [源单位]、eUnit 源单位枚举、fTankHeight 罐内有效高度 [m]；fOut 折算结果 [m]；
        返回 TRUE 表示 fOut 可信。% 通道要求 fTankHeight > 0，否则判不可信（不除零）。
  边界：① 除零防护：仅对 100 常量做除法，罐高为 0 时 % 通道直接判不可信；② 未知枚举 / 非有限输入 → FALSE + 0.0；
        ③ 三个浮点入参逐一做非有限闸；零全局、零物理地址、零库件依赖。
*)

(*-----------------------------------------------------------------------------
 * 枚举: E_DL_LvlUnit（液位单位，归属本文件，全库唯一定义）
 *----------------------------------------------------------------------------*)
TYPE E_DL_LvlUnit :
(
    eMeter    := 0,    // 米（基准单位） [m] / Metre, the base unit
    eMilliMeter := 1,  // 毫米 [mm] / Millimetre
    ePercent  := 2     // 百分比（按罐高折算） [%] / Percent of the tank height
);
END_TYPE

FUNCTION FC_DL_LevelUnitConvert : BOOL
VAR_INPUT
    fIn        : LREAL := 0.0;         // 输入值 [源单位] / The input value in the source unit
    eUnit      : E_DL_LvlUnit;         // 源单位枚举 [—] / The source unit enumeration
    fTankHeight : LREAL := 1.0;        // 罐内有效高度（% 通道必需 > 0） [m] / The effective tank height for percent
END_VAR
VAR_OUTPUT
    fOut : LREAL;                      // 折算结果 [m] / The converted value in the base unit
END_VAR
VAR CONSTANT
    DL_LV_MM   : LREAL := 0.001;       // 1 mm 折 m 的系数 [-] / millimetre to metre
    DL_LV_HUND : LREAL := 100.0;       // 百分比满量程分母 [-] / The percent full scale divisor
    DL_LV_INF  : LREAL := 1.0E30;      // 非有限 / 越界判据上限 [-] / The magnitude gate
    DL_LV_EPS  : LREAL := 1.0E-9;      // 罐高判零容差 [-] / The tank height zero tolerance
    DL_LV_Z    : LREAL := 0.0;         // 浮点零常量 [m] / The floating point zero constant
END_VAR

FC_DL_LevelUnitConvert := FALSE;                          // 返回值预置假 / preset the return false
fOut := DL_LV_Z;                                          // 输出预置零哨兵 [m] / preset the zero sentinel
IF (fIn <> fIn) OR (ABS(fIn) > DL_LV_INF) THEN            // 输入自反判 NaN 或越限判 Inf / the input gate
    fOut := DL_LV_Z;                                      // 非有限值输出零哨兵 [m] / zero the non finite input
ELSIF (fTankHeight <> fTankHeight) OR (ABS(fTankHeight) > DL_LV_INF) THEN // 罐高非有限闸 / the tank height gate
    fOut := DL_LV_Z;                                      // 罐高非法输出零哨兵 [m] / zero sentinel on an invalid height
ELSE
    CASE eUnit OF
        E_DL_LvlUnit.eMeter:                              // 基准单位直通 / the base unit passes through
            fOut := fIn;                                  // 直通不换算 [m] / pass through unchanged
            FC_DL_LevelUnitConvert := TRUE;               // 结果可信 / the result is valid
        E_DL_LvlUnit.eMilliMeter:                         // 毫米折米 / millimetre to metre
            fOut := fIn * DL_LV_MM;                       // 乘 0.001 [m] / multiply by the factor
            FC_DL_LevelUnitConvert := TRUE;               // 结果可信 / the result is valid
        E_DL_LvlUnit.ePercent:                            // 百分比按罐高折算 / percent of the tank height
            IF (fTankHeight > DL_LV_EPS) THEN             // 罐高为正才可折算（除零防护） / a positive height is required
                fOut := (fIn / DL_LV_HUND) * fTankHeight; // 先除常量 100 再乘罐高 [m] / divide then multiply
                FC_DL_LevelUnitConvert := TRUE;           // 结果可信 / the result is valid
            ELSE
                fOut := DL_LV_Z;                          // 罐高为零输出零哨兵 [m] / zero sentinel on a zero height
                FC_DL_LevelUnitConvert := FALSE;          // 不可信 / not valid
            END_IF
    ELSE
        fOut := DL_LV_Z;                                  // 未知枚举输出零哨兵 [m] / zero sentinel on an unknown unit
        FC_DL_LevelUnitConvert := FALSE;                  // 未知枚举不可信 / an unknown unit is not valid
    END_CASE
END_IF
END_FUNCTION

(* ---- FC_DL_MapRangePercent.st ---- *)
(*
  FC_DL_MapRangePercent —— 百分比与工程值互映，枚举方向
  分类：DL_Base | 复杂度：1 | 轮次：R86
  开源溯源：道莅原创（clean-room 自研，纯 IEC 61131-3 通用算法），无外部代码引用
  许可证：MIT
  职责：按 eDir 方向做百分比与工程值互映：
        ePctToEng：fIn 视为百分比 0..100，映射到 [fOutMin, fOutMax]；
        eEngToPct：fIn 视为工程量，映射到百分比 0..100（先钳到量程）。
  契约：fIn 输入值、eDir 方向枚举、fEngMin/fEngMax 工程量程端点；fOut 结果 [目标单位]；返回 TRUE 表示可信。
  边界：① 量程退化校验（容差 DL_MP_EPS）；② 除零防护：分母先过退化闸；③ 浮点入参逐一非有限闸；
        ④ CASE 含 ELSE 兜底拦非法方向；零全局、零物理地址、零库件依赖。
*)

(*-----------------------------------------------------------------------------
 * 枚举: E_DL_MapDir（映射方向，归属本文件，全库唯一定义）
 *----------------------------------------------------------------------------*)
TYPE E_DL_MapDir :
(
    ePctToEng := 0,    // 百分比 → 工程值 [—] / Percent to engineering value
    eEngToPct := 1     // 工程值 → 百分比 [—] / Engineering value to percent
);
END_TYPE

FUNCTION FC_DL_MapRangePercent : BOOL
VAR_INPUT
    fIn     : LREAL := 0.0;            // 输入值 [源单位] / The input value in the source unit
    eDir    : E_DL_MapDir;             // 映射方向枚举 [—] / The mapping direction
    fEngMin : LREAL := 0.0;            // 工程量程下端点 [工程单位] / The engineering range low end
    fEngMax : LREAL := 100.0;          // 工程量程上端点 [工程单位] / The engineering range high end
END_VAR
VAR_OUTPUT
    fOut : LREAL;                      // 结果 [目标单位] / The result in the target unit
END_VAR
VAR
    xBad     : BOOL;                   // 参数非法标志 [—] / The parameter invalid flag
    fInClamp : LREAL;                  // 钳位后的输入 [源单位] / The clamped input value
    fEngSpan : LREAL;                  // 工程量程跨度 [工程单位] / The engineering span
END_VAR
VAR CONSTANT
    DL_MP_EPS   : LREAL := 1.0E-9;     // 浮点比较容差 [-] / The floating point comparison tolerance
    DL_MP_INF   : LREAL := 1.0E30;     // 非有限 / 越界判据上限 [-] / The magnitude gate
    DL_MP_Z     : LREAL := 0.0;        // 浮点零常量 [-] / The floating point zero constant
    DL_MP_HUND  : LREAL := 100.0;      // 百分比满量程 [-] / The percent full scale
END_VAR

FC_DL_MapRangePercent := FALSE;                           // 返回值预置假 / preset the return false
fOut := DL_MP_Z;                                          // 输出预置零哨兵 / preset the zero sentinel
xBad := FALSE;                                            // 非法标志预置假 / preset the invalid flag false
IF (fIn <> fIn) OR (ABS(fIn) > DL_MP_INF) THEN            // 输入非有限闸 / the input gate
    xBad := TRUE;                                         // 置非法标志 / raise the invalid flag
END_IF
IF (fEngMin <> fEngMin) OR (ABS(fEngMin) > DL_MP_INF) THEN // 工程下端非有限闸 / the engineering low end gate
    xBad := TRUE;                                         // 置非法标志 / raise the invalid flag
END_IF
IF (fEngMax <> fEngMax) OR (ABS(fEngMax) > DL_MP_INF) THEN // 工程上端非有限闸 / the engineering high end gate
    xBad := TRUE;                                         // 置非法标志 / raise the invalid flag
END_IF
fEngSpan := fEngMax - fEngMin;                            // 工程量程跨度 [工程单位] / the engineering span
IF ABS(fEngSpan) < DL_MP_EPS THEN                         // 量程退化（除零防护） / the degenerate span
    xBad := TRUE;                                         // 置非法标志 / raise the invalid flag
END_IF
IF NOT xBad THEN                                          // 参数全通过才映射 / map only when all parameters pass
    CASE eDir OF
        E_DL_MapDir.ePctToEng:                            // 百分比转工程值 / percent to engineering value
            fInClamp := fIn;                              // 输入接管 [%] / take the input value
            IF fInClamp < DL_MP_Z THEN                    // 百分比低于零 / below zero percent
                fInClamp := DL_MP_Z;                      // 钳到零 [%] / clamp to zero
            END_IF
            IF fInClamp > DL_MP_HUND THEN                 // 百分比高于一百 / above one hundred percent
                fInClamp := DL_MP_HUND;                   // 钳到一百 [%] / clamp to one hundred
            END_IF
            fOut := fEngMin + (fInClamp / DL_MP_HUND) * fEngSpan; // 线性换算（除常量） [工程单位] / the conversion
            FC_DL_MapRangePercent := TRUE;                // 结果可信 / the result is valid
        E_DL_MapDir.eEngToPct:                            // 工程值转百分比 / engineering value to percent
            fInClamp := fIn;                              // 输入接管 [工程单位] / take the input value
            IF fEngSpan > DL_MP_Z THEN                    // 正常量程方向 / the normal span direction
                IF fInClamp < fEngMin THEN                // 低于下端点 / below the low end
                    fInClamp := fEngMin;                  // 钳到下端点 [工程单位] / clamp to the low end
                END_IF
                IF fInClamp > fEngMax THEN                // 高于上端点 / above the high end
                    fInClamp := fEngMax;                  // 钳到上端点 [工程单位] / clamp to the high end
                END_IF
            ELSE                                          // 反向量程 / the reversed span
                IF fInClamp > fEngMin THEN                // 高于下端（反向即越小越远） / above the low end
                    fInClamp := fEngMin;                  // 钳到下端点 [工程单位] / clamp to the low end
                END_IF
                IF fInClamp < fEngMax THEN                // 低于上端点 / below the high end
                    fInClamp := fEngMax;                  // 钳到上端点 [工程单位] / clamp to the high end
                END_IF
            END_IF
            fOut := ((fInClamp - fEngMin) / fEngSpan) * DL_MP_HUND; // 反向换算（分母已证非零） [%] / the conversion
            FC_DL_MapRangePercent := TRUE;                // 结果可信 / the result is valid
    ELSE
        fOut := DL_MP_Z;                                  // 非法方向输出零哨兵 / zero sentinel on an illegal direction
        FC_DL_MapRangePercent := FALSE;                   // 非法方向不可信 / an illegal direction is not valid
    END_CASE
END_IF
END_FUNCTION

(* ---- FC_DL_SaturateAdd.st ---- *)
(*
  FC_DL_SaturateAdd  —  饱和加减运算 / Saturating add and subtract
  分类 Category : DL_Base
  码位 Code     : 16#01_0_00
  版本 Version  : 1.0.0
  来源 Source   : t2-1-lgf-math — IEC 61131-3 标准语义的道莅防御性实现
  溯源 Origin   : clean-room 实现，通用饱和算术语义，未复制任何源码行
  功能 Function : 1) 以 LINT 宽域中间量计算 nInA ± nInB（Add/Sub 两模式），杜绝 DINT 先加后判的回绕静默翻号；
                  2) 结果先与 [nLimitLo, nLimitHi] 组态区间钳制，再与 DINT 可表达域钳制，输出最终 nOut；
                  3) bClamped 指示本调用发生了钳制（每调用无条件重算，无锁存）。
  边界 Boundary : ① nLimitLo > nLimitHi 判组态错置码，输出 nLimitLo（安全侧下界）且 bClamped := TRUE；
                  ② 结果超出 DINT 可表达域时饱和到对应 DINT 极限并 bClamped := TRUE（DINT ± DINT 在 LINT 内必不溢出，此分支为防御性兜底）；
                  ③ eOp 落入未知值由 CASE ELSE 拦截：置码、输出 0、bClamped := TRUE（不猜运算方向）；
                  ④ 解除式自证：bClamped 为每调用重算量，下一调用结果重新落入区间即自动解除（无 bReset、无锁存）；
                  ⑤ 本件为纯函数：无 VAR 记忆量、无定时器、无边沿实例，可离平台编译。
  依赖 Depends  : 仅 Standard.library（无库调用）；枚举 E_DL_SatOp 随本件发布
  码表 Error codes（本件格 01_0_00，子码步进 +0x100）:
    16#0001_0100 信息级：结果被钳制（bClamped = TRUE，不置故障）
    16#0001_0200 故障级：组态非法 nLimitLo > nLimitHi，输出安全侧下界
    16#0001_0300 故障级：运算模式 eOp 非法（CASE ELSE 兜底）

  修订历史 Revision :
    2026-11-18  v1.0.0  R38 首版
*)

TYPE E_DL_SatOp :
(
    eAdd := 0,   // 加法模式 / Addition mode
    eSub := 1    // 减法模式 / Subtraction mode
);
END_TYPE

FUNCTION FC_DL_SaturateAdd : BOOL
VAR_INPUT
    nInA     : DINT;                 // 操作数 A / Operand A
    nInB     : DINT;                 // 操作数 B / Operand B
    eOp      : E_DL_SatOp;           // 运算模式（Add/Sub）/ Operation mode, Add or Sub
    nLimitHi : DINT;                 // 组态上限 [DINT] / Configured upper limit
    nLimitLo : DINT;                 // 组态下限 [DINT] / Configured lower limit
END_VAR
VAR_OUTPUT
    nOut     : DINT;                 // 钳制后结果 / Saturated result
    bClamped : BOOL;                 // 本调用发生钳制 / Clamped on this call, recomputed per call
    nErrId   : UDINT;                // 事件码，0 = 无事件 / Event code, 0 = none
END_VAR
VAR
    liWork : LINT;                  // 宽域中间量（FC 局部临时量，每调用重算，非记忆量）/ Wide scratch, temp per call
END_VAR
VAR CONSTANT
    DL_DINT_HI : LINT := 2147483647;   // DINT 可表达上界 / Expressible DINT upper bound
    DL_DINT_LO : LINT := -2147483648;  // DINT 可表达下界 / Expressible DINT lower bound
END_VAR

(* —— 段 1：单拍量缺省与组态闸（纯函数，每调用重算） —— *)
nOut     := 0;                        // 输出缺省 0
bClamped := FALSE;                    // 钳制标志每调用重算（无锁存，解除式自证）
nErrId   := 16#0000_0000;             // 事件码缺省无事件

IF nLimitLo > nLimitHi THEN
    nOut     := nLimitLo;             // 组态错：输出安全侧下界（规格强制）
    bClamped := TRUE;                 // 组态错视为钳制
    nErrId   := 16#0001_0200;         // 故障级：组态非法
    FC_DL_SaturateAdd := FALSE;       // 返回值：运算未受理
    RETURN;                            // 组态非法不进入运算
END_IF

(* —— 段 2：LINT 宽域运算（禁先 DINT 相加再判溢出） —— *)
CASE eOp OF

E_DL_SatOp.eAdd:
    liWork := LINT(nInA) + LINT(nInB);   // 宽域加法，DINT±DINT 必不溢出 LINT
    FC_DL_SaturateAdd := TRUE;           // 运算已受理

E_DL_SatOp.eSub:
    liWork := LINT(nInA) - LINT(nInB);   // 宽域减法
    FC_DL_SaturateAdd := TRUE;           // 运算已受理

ELSE
    nOut   := 0;                    // 未知模式：输出 0（不猜方向）
    bClamped := TRUE;               // 视为异常钳制
    nErrId := 16#0001_0300;         // 故障级：运算模式非法
    FC_DL_SaturateAdd := FALSE;     // 运算未受理
    RETURN;

END_CASE

(* —— 段 3：先 DINT 可表达域钳制，再组态区间钳制（顺序不可倒置） —— *)
IF liWork > DL_DINT_HI THEN
    liWork   := DL_DINT_HI;         // 超上界：饱和到 DINT 上限
    bClamped := TRUE;               // 钳制标志
    nErrId   := 16#0001_0100;       // 信息级：结果被钳制
ELSIF liWork < DL_DINT_LO THEN
    liWork   := DL_DINT_LO;         // 超下界：饱和到 DINT 下限
    bClamped := TRUE;
    nErrId   := 16#0001_0100;       // 信息级：结果被钳制
END_IF

IF liWork > LINT(nLimitHi) THEN
    liWork   := LINT(nLimitHi);     // 超组态上限：钳到上限
    bClamped := TRUE;
    nErrId   := 16#0001_0100;       // 信息级：结果被钳制
ELSIF liWork < LINT(nLimitLo) THEN
    liWork   := LINT(nLimitLo);     // 低于组态下限：钳到下限
    bClamped := TRUE;
    nErrId   := 16#0001_0100;       // 信息级：结果被钳制
END_IF

(* —— 段 4：出口单点映射 —— *)
nOut := DINT(liWork);               // 宽域结果回落 DINT（已经两段钳制，必在表达域内）

END_FUNCTION

(* ---- FC_DL_SpecificHeatUnitConvert.st ---- *)
(*
  FC_DL_SpecificHeatUnitConvert —— 比热容换算 kJ/(kg*K) 与 BTU/(lb*F)
  分类：DL_Base | 复杂度：1 | 轮次：R86
  开源溯源：道莅原创（clean-room 自研，纯 IEC 61131-3 通用算法），无外部代码引用
  许可证：MIT
  职责：把比热容统一折算到基准单位 kJ/(kg*K)（1 BTU/(lb*F) = 4.1868 kJ/(kg*K)）。
  契约：fIn 输入值 [源单位]，eUnit 源单位枚举；fOut 折算结果 [kJ/(kg*K)]；返回 TRUE 表示 fOut 可信。
  边界：未知枚举 / 非有限输入 → 返回 FALSE，fOut 给 0.0 哨兵；无除法，零全局、零物理地址、零库件依赖。
*)

(*-----------------------------------------------------------------------------
 * 枚举: E_DL_ShcUnit（比热容单位，归属本文件，全库唯一定义）
 *----------------------------------------------------------------------------*)
TYPE E_DL_ShcUnit :
(
    eKjPerKgK  := 0,   // 千焦每千克开（基准单位） [kJ/(kg*K)] / Kilojoule per kilogram kelvin, the base unit
    eBtuPerLbF := 1    // 英热单位每磅华氏度 [BTU/(lb*F)] / British thermal unit per pound fahrenheit
);
END_TYPE

FUNCTION FC_DL_SpecificHeatUnitConvert : BOOL
VAR_INPUT
    fIn   : LREAL := 0.0;              // 输入值 [源单位] / The input value in the source unit
    eUnit : E_DL_ShcUnit;              // 源单位枚举 [—] / The source unit enumeration
END_VAR
VAR_OUTPUT
    fOut : LREAL;                      // 折算结果 [kJ/(kg*K)] / The converted value in the base unit
END_VAR
VAR CONSTANT
    DL_SC_BTU : LREAL := 4.1868;       // 1 BTU/(lb*F) 折 kJ/(kg*K) 的系数 [-] / BTU per lb F to kJ per kg K
    DL_SC_INF : LREAL := 1.0E30;       // 非有限 / 越界判据上限 [-] / The magnitude gate
    DL_SC_Z   : LREAL := 0.0;          // 浮点零常量 [kJ/(kg*K)] / The floating point zero constant
END_VAR

FC_DL_SpecificHeatUnitConvert := FALSE;                   // 返回值预置假 / preset the return false
fOut := DL_SC_Z;                                          // 输出预置零哨兵 [kJ/(kg*K)] / preset the zero sentinel
IF (fIn <> fIn) OR (ABS(fIn) > DL_SC_INF) THEN            // 自反判 NaN 或越限判 Inf / NaN or Inf
    fOut := DL_SC_Z;                                      // 非有限值输出零哨兵 [kJ/(kg*K)] / zero the non finite input
ELSE
    CASE eUnit OF
        E_DL_ShcUnit.eKjPerKgK:                           // 基准单位直通 / the base unit passes through
            fOut := fIn;                                  // 直通不换算 [kJ/(kg*K)] / pass through unchanged
            FC_DL_SpecificHeatUnitConvert := TRUE;        // 结果可信 / the result is valid
        E_DL_ShcUnit.eBtuPerLbF:                          // 英热单位每磅华氏度 / BTU per pound fahrenheit
            fOut := fIn * DL_SC_BTU;                      // 乘 4.1868 [kJ/(kg*K)] / multiply by the factor
            FC_DL_SpecificHeatUnitConvert := TRUE;        // 结果可信 / the result is valid
    ELSE
        fOut := DL_SC_Z;                                  // 未知枚举输出零哨兵 [kJ/(kg*K)] / zero sentinel on an unknown unit
        FC_DL_SpecificHeatUnitConvert := FALSE;           // 未知枚举不可信 / an unknown unit is not valid
    END_CASE
END_IF
END_FUNCTION

(* ---- FC_DL_StringCompareNatural.st ---- *)
(*==============================================================================
 * 组件名称 (Component)  : FC_DL_StringCompareNatural
 * 所属子库 (Sublibrary) : DL_Base
 * 当前版本 (Version)    : 1.0.0
 * 兼容性   (Platform)   : CODESYS 3.5+ / TwinCAT 3 / 汇川 InoProShop / 施耐德 Machine Expert
 *                         仅依赖 IEC 61131-3 标准字符串九函数（LEN / MID / LEFT / CONCAT / DELETE / FIND），零厂商私有库
 * 功能描述 (Function)   : 自然序比较（Human sort / natural sort）。规则：
 *                           · 双方同位置均为数字时，各自提取完整数字段，按「数值」比较
 *                             （去前导零后先比位数、同位数再逐位比较），故 A2 < A10；
 *                           · 其余位置按单字符序数比较，序数由排序字符集常量
 *                             DL_SCN_ORDER 的 FIND 位置给出（集合外字符序数记 0，排最前）；
 *                           · 公共前缀耗尽后，剩余字符多者更大（A < AB）。
 *                         全程用 FIND(集合, 单字符) 取序数，不依赖平台字符串比较运算符或
 *                         字符码强转方言（R3 纯标准函数路径）。
 * 接口     (Interface)  : 输入 sInA 左串、sInB 右串 [-]；
 *                         输出 iResult 比较结果（-1 左小 / 0 相等 / 1 左大）[-]、
 *                         bEqual 是否相等、eErrCode 错误码（E_DL_StrNatErr）；
 *                         返回值 = bValid 比较可信标志（TRUE = iResult 可信）。
 * 边界     (Boundary)   : ① 属主边界：只做比较，不做排序（排序归调用方的数组管理）、
 *                         不做大小写折叠（'A' 与 'a' 序数不同，A 在前）。
 *                         ② 数字段归一：去前导零后 '007' 与 '7' 相等（数值 7），
 *                         故 "A007" = "A7"（iResult=0）；长度差由去零后的位数决定。
 *                         ③ 序数集合只含 0-9 / A-Z / a-z；标点与空格序数记 0（同序则继续后移，
 *                         不判等、不报错），排序稳定性由调用方的稳定排序保证。
 *                         ④ 长度均钳位至 255（缓冲可表性），双向扫描严格有界。
 *                         ⑤ 内层数字段提取循环亦以上界 _udLenA/_udLenB 收口，无越界。
 *                         ⑥ 零全局耦合（无 GVL / VAR_EXTERNAL / 物理地址）。
 * 分工声明 (Scope)      : 与 `FC_DL_StringReverse` 分工：位序重排归那件、序比较归本件；
 *                         与 `FC_DL_StringIsNumeric` 分工：整串数值判定归那件。
 * 来源标签 (Source Tag) : 原创实现（无外部代码引入）
 * 码表     (Codes)      : 本件不占用全局数字码位；出口为 BOOL + INT + BOOL +
 *                         本文件内定义 enum E_DL_StrNatErr（全库唯一）。
 * 红线自检 (Redline)    : R1 ✓ 零 GVL/VAR_EXTERNAL ｜ R2 ✓ 零 %I/%Q/%M ｜ R3 ✓ 纯 IEC 61131-3
 *                         R4 ✓ 双层循环上界收口 + 去前导零守恒 + 序数集合法（无字符码强转） ｜ R5 ✓ 声明逐行同行双语注释
 *                         R6 N/A（纯函数无状态机） ｜ R7 N/A（无实例调用）
 * 修订历史 (Revision)   : 2026-11-23  v1.0.0  R77 首版（批次 B2 · 序号 9）
 * 验收向量 (Acceptance) : ① sInA='A2', sInB='A10' → iResult=-1（数字段 2 < 10）, bEqual=FALSE, eOk；
 *                         ② sInA='A2', sInB='A2' → iResult=0, bEqual=TRUE；
 *                         ③ sInA='A007', sInB='A7' → 去零后数值相同 → iResult=0, bEqual=TRUE；
 *                         ④ sInA='A', sInB='AB' → 公共前缀耗尽，右串剩余 → iResult=-1；
 *                         ⑤ sInA='B1', sInB='A99' → 首字符序数 B > A → iResult=1；
 *                         ⑥ sInA='', sInB='' → iResult=0, bEqual=TRUE, eOk。
 *==============================================================================*)

(*-----------------------------------------------------------------------------
 * 枚举: E_DL_StrNatErr（自然序比较错误码，归属 DL_Base，与本件同文件，全库唯一属主）
 *----------------------------------------------------------------------------*)
TYPE E_DL_StrNatErr :
(
    eOk      := 0,   // 信息级：比较完成，结果可信 / Info: comparison completed, result trustworthy
    eClampLen:= 1    // 信息级：输入超缓冲上限已按 255 字符比较 / Info: inputs clamped to 255 chars for comparison
);
END_TYPE

FUNCTION FC_DL_StringCompareNatural : BOOL
VAR_INPUT
    sInA : STRING(255);   // 左串 [-] / Left string
    sInB : STRING(255);   // 右串 [-] / Right string
END_VAR
VAR_OUTPUT
    iResult : INT;        // 比较结果：-1 左小 / 0 相等 / 1 左大 [-] / Compare result: -1 less, 0 equal, 1 greater
    bEqual  : BOOL;       // 是否相等（iResult=0） [-] / Whether equal, iResult equals zero
    eErrCode: E_DL_StrNatErr; // 错误码出口 [-] / Error code outlet
END_VAR
VAR
    _udLenA  : UDINT;       // 左串生效长度 [字符] / Effective left length [chars]
    _udLenB  : UDINT;       // 右串生效长度 [字符] / Effective right length [chars]
    _udA     : UDINT;       // 左串游标（1 基） [-] / Left cursor, 1-based
    _udB     : UDINT;       // 右串游标（1 基） [-] / Right cursor, 1-based
    _udKa    : UDINT;       // 数字段内位序 [-] / Bit index inside digit run
    _udRunA  : UDINT;       // 左数字段长度 [字符] / Left digit run length [chars]
    _udRunB  : UDINT;       // 右数字段长度 [字符] / Right digit run length [chars]
    _rkA     : UDINT;       // 左字符序数（0 = 集合外） [-] / Left character rank, 0 means outside set
    _rkB     : UDINT;       // 右字符序数（0 = 集合外） [-] / Right character rank, 0 means outside set
    _sChA    : STRING(255); // 左串当前单字符 [-] / Current left character
    _sChB    : STRING(255); // 右串当前单字符 [-] / Current right character
    _sRunA   : STRING(255); // 左数字段（已去前导零） [-] / Left digit run, leading zeros stripped
    _sRunB   : STRING(255); // 右数字段（已去前导零） [-] / Right digit run, leading zeros stripped
    _iRes    : INT;         // 比较结果内部累加 [-] / Internal compare result
END_VAR
VAR CONSTANT
    DL_SCN_SET_DIGIT : STRING(255) := '0123456789';   // 数字字符集 [-] / Digit character set
    DL_SCN_SET_ZERO  : STRING(255) := '0';            // 零字符集（去前导零用） [-] / Zero character set for leading-zero strip
    DL_SCN_ORDER     : STRING(255) := '0123456789ABCDEFGHIJKLMNOPQRSTUVWXYZabcdefghijklmnopqrstuvwxyz'; // 序数字符集 [-] / Rank character set
    DL_SCN_LEN_MAX   : UINT := 255;                   // 缓冲上限（STRING(255) 契约） [字符] / Buffer ceiling [chars]
    DL_SCN_START     : UDINT := 1;                    // 字符串起始位置（IEC 1 基） [-] / String start position, 1-based
    DL_SCN_ONE_LEN   : UDINT := 1;                    // 单字符长度常量 [字符] / Single character length constant
    DL_SCN_HIT_ONE   : UDINT := 1;                    // FIND 首位命中的比较值 [-] / Compare value for first-position hit
END_VAR

(* —— 段 0：出口预置安全值 —— *)
FC_DL_StringCompareNatural := FALSE;               // 返回值预置不可信 / Return preset untrustworthy
iResult  := 0;                                     // 比较结果哨兵：相等 / Result sentinel: equal
bEqual   := FALSE;                                 // 相等标志预置否 / Equality flag preset false
eErrCode := E_DL_StrNatErr.eClampLen;              // 预置最严码（本件仅信息级码） / Preset strictest code

(* —— 段 1：长度实测与上域钳位（双向扫描严格有界） —— *)
_udLenA := LEN(sInA);                              // 左串字符数 / Left length
_udLenB := LEN(sInB);                              // 右串字符数 / Right length
IF (_udLenA > UINT_TO_UDINT(DL_SCN_LEN_MAX)) OR (_udLenB > UINT_TO_UDINT(DL_SCN_LEN_MAX)) THEN
    eErrCode := E_DL_StrNatErr.eClampLen;          // 信息级钳位码 / Info clamp code
ELSE
    eErrCode := E_DL_StrNatErr.eOk;                // 信息级成功预置 / Info success preset
END_IF
IF _udLenA > UINT_TO_UDINT(DL_SCN_LEN_MAX) THEN
    _udLenA := UINT_TO_UDINT(DL_SCN_LEN_MAX);      // 左串钳位 / Left clamped
END_IF
IF _udLenB > UINT_TO_UDINT(DL_SCN_LEN_MAX) THEN
    _udLenB := UINT_TO_UDINT(DL_SCN_LEN_MAX);      // 右串钳位 / Right clamped
END_IF

(* —— 段 2：游标与结果预清零（不含保持量，逐次比较独立） —— *)
_udA  := DL_SCN_START;
_udB  := DL_SCN_START;
_iRes := 0;

(* —— 段 3：主扫描（双游标均在界内且尚未分出胜负） —— *)
WHILE (_udA <= _udLenA) AND (_udB <= _udLenB) AND (_iRes = 0) DO
    _sChA := MID(sInA, DL_SCN_ONE_LEN, _udA);      // 取左串当前字符 / Take left current character
    _sChB := MID(sInB, DL_SCN_ONE_LEN, _udB);      // 取右串当前字符 / Take right current character

    IF (FIND(DL_SCN_SET_DIGIT, _sChA) > 0) AND (FIND(DL_SCN_SET_DIGIT, _sChB) > 0) THEN
        (* —— 段 3a：双方均为数字 → 提取完整数字段按数值比较 —— *)
        _sRunA := '';                              // 左数字段清空 / Clear left run
        WHILE (_udA <= _udLenA) AND (FIND(DL_SCN_SET_DIGIT, MID(sInA, DL_SCN_ONE_LEN, _udA)) > 0) DO
            _sRunA := CONCAT(_sRunA, MID(sInA, DL_SCN_ONE_LEN, _udA));   // 逐位累积左数字段 / Accumulate left digit
            _udA   := _udA + 1;                    // 游标越过该位 / Cursor passes this digit
        END_WHILE
        _sRunB := '';                              // 右数字段清空 / Clear right run
        WHILE (_udB <= _udLenB) AND (FIND(DL_SCN_SET_DIGIT, MID(sInB, DL_SCN_ONE_LEN, _udB)) > 0) DO
            _sRunB := CONCAT(_sRunB, MID(sInB, DL_SCN_ONE_LEN, _udB));   // 逐位累积右数字段 / Accumulate right digit
            _udB   := _udB + 1;
        END_WHILE

        (* 去前导零：保留至少一位（"000" 归一为 "0"） *)
        WHILE (LEN(_sRunA) > DL_SCN_ONE_LEN) AND (FIND(DL_SCN_SET_ZERO, LEFT(_sRunA, DL_SCN_ONE_LEN)) = DL_SCN_HIT_ONE) DO
            _sRunA := DELETE(_sRunA, DL_SCN_ONE_LEN, DL_SCN_START);      // 删首零 / Delete leading zero
        END_WHILE
        WHILE (LEN(_sRunB) > DL_SCN_ONE_LEN) AND (FIND(DL_SCN_SET_ZERO, LEFT(_sRunB, DL_SCN_ONE_LEN)) = DL_SCN_HIT_ONE) DO
            _sRunB := DELETE(_sRunB, DL_SCN_ONE_LEN, DL_SCN_START);      // 删首零 / Delete leading zero
        END_WHILE

        _udRunA := LEN(_sRunA);                    // 左段位数 / Left digit count
        _udRunB := LEN(_sRunB);                    // 右段位数 / Right digit count
        IF _udRunA < _udRunB THEN
            _iRes := -1;                           // 位数少者数值小 / Fewer digits is smaller
        ELSIF _udRunA > _udRunB THEN
            _iRes := 1;                            // 位数多者数值大 / More digits is greater
        ELSE
            _udKa := DL_SCN_START;                 // 同位数逐位比较 / Same digit count: compare per digit
            WHILE (_udKa <= _udRunA) AND (_iRes = 0) DO
                _rkA := FIND(DL_SCN_SET_DIGIT, MID(_sRunA, DL_SCN_ONE_LEN, _udKa));  // 左位序数 / Left digit rank
                _rkB := FIND(DL_SCN_SET_DIGIT, MID(_sRunB, DL_SCN_ONE_LEN, _udKa));  // 右位序数 / Right digit rank
                IF _rkA < _rkB THEN
                    _iRes := -1;                   // 左位小 / Left digit smaller
                ELSIF _rkA > _rkB THEN
                    _iRes := 1;                    // 左位大 / Left digit greater
                END_IF
                _udKa := _udKa + 1;                // 位序步进 / Advance digit index
            END_WHILE
        END_IF
    ELSE
        (* —— 段 3b：非数字段 → 按字符序数比较 —— *)
        _rkA := FIND(DL_SCN_ORDER, _sChA);         // 左字符序数（集合外 = 0） / Left rank, outside set is zero
        _rkB := FIND(DL_SCN_ORDER, _sChB);         // 右字符序数（集合外 = 0） / Right rank, outside set is zero
        IF _rkA < _rkB THEN
            _iRes := -1;                           // 左字符序数小 / Left character rank smaller
        ELSIF _rkA > _rkB THEN
            _iRes := 1;                            // 左字符序数大 / Left character rank greater
        END_IF
        _udA := _udA + 1;                          // 双游标同步步进 / Advance both cursors
        _udB := _udB + 1;
    END_IF
END_WHILE

(* —— 段 4：公共前缀耗尽后的长度裁决（剩余字符多者更大） —— *)
IF _iRes = 0 THEN
    IF _udA <= _udLenA THEN
        _iRes := 1;                                // 左串有剩余 → 左大 / Left has remainder: greater
    ELSIF _udB <= _udLenB THEN
        _iRes := -1;                               // 右串有剩余 → 左小 / Right has remainder: less
    ELSE
        _iRes := 0;                                // 同时耗尽 → 相等 / Both exhausted: equal
    END_IF
END_IF

(* —— 段 5：导出结果与相等标志 —— *)
iResult := _iRes;                                  // 导出比较结果 / Export compare result
bEqual  := (_iRes = 0);                            // 相等标志 / Equality flag
FC_DL_StringCompareNatural := TRUE;                // 比较可信 / Comparison trustworthy

END_FUNCTION

(* ---- FC_DL_StringCountChar.st ---- *)
(*==============================================================================
 * 组件名称 (Component)  : FC_DL_StringCountChar
 * 所属子库 (Sublibrary) : DL_Base
 * 当前版本 (Version)    : 1.0.0
 * 兼容性   (Platform)   : CODESYS 3.5+ / TwinCAT 3 / 汇川 InoProShop / 施耐德 Machine Expert
 *                         仅依赖 IEC 61131-3 标准字符串九函数（LEN / LEFT / MID / FIND），零厂商私有库
 * 功能描述 (Function)   : 统计指定字符在字符串中的出现次数。典型用途：HMI 报文
 *                         分隔符计数（判断字段数 = 分隔符数 + 1）、协议帧结构预校验。
 *                         逐字符扫描，用 FIND(单字符, 实测单字符) = 1 做单字符等值判定
 *                         （纯 IEC 标准函数路径，不依赖平台 STRING 比较运算符方言；
 *                         单字符串 A 与 B 相等 ⇔ FIND(A,B)=1）。
 *                         填充字符取 sChar 首字符，故传入多字符串时按首字符计。
 * 接口     (Interface)  : 输入 sIn 被扫描字符串 [-]、sChar 目标字符（取首字符）[-]；
 *                         输出 uiCount 出现次数 [次]、uiLen 扫描字符数 [字符]、
 *                         eErrCode 错误码（E_DL_StrCountErr）；
 *                         返回值 = bValid 统计可信标志（TRUE = uiCount 可信）。
 * 边界     (Boundary)   : ① 属主边界：只统计单字符，不做多字符串（子串）计数、
 *                         不做分隔符拆分（拆分归 FC_DL_StringSplitPair）。
 *                         ② sChar 为空串 → 故障级 eEmptyChar，uiCount 哨兵 0。
 *                         ③ sIn 为空串 → 合法，uiCount=0、uiLen=0、eOk（空串零命中）。
 *                         ④ 扫描上界取 uiLen（<=255），循环严格有界，无越界读取。
 *                         ⑤ 零全局耦合（无 GVL / VAR_EXTERNAL / 物理地址）。
 * 分工声明 (Scope)      : 与 `FC_DL_StringSplitPair` 分工：本件只计数不拆分；
 *                         与 `FC_DL_StringRemoveWhitespace` 分工：空白剔除归那件。
 * 来源标签 (Source Tag) : 原创实现（无外部代码引入）
 * 码表     (Codes)      : 本件不占用全局数字码位；出口为 BOOL + UINT +
 *                         本文件内定义 enum E_DL_StrCountErr（全库唯一）。
 * 红线自检 (Redline)    : R1 ✓ 零 GVL/VAR_EXTERNAL ｜ R2 ✓ 零 %I/%Q/%M ｜ R3 ✓ 纯 IEC 61131-3
 *                         R4 ✓ 空字符域闸 + 扫描上界钳位 + 单字符等值判定 ｜ R5 ✓ 声明逐行同行双语注释
 *                         R6 N/A（纯函数无状态机） ｜ R7 N/A（无实例调用）
 * 修订历史 (Revision)   : 2026-11-23  v1.0.0  R77 首版（批次 B2 · 序号 3）
 * 验收向量 (Acceptance) : ① sIn='A,B,C,D', sChar=',' → uiCount=3, uiLen=7, eOk, TRUE；
 *                         ② sIn='ABCD', sChar=',' → uiCount=0, uiLen=4, eOk, TRUE；
 *                         ③ sIn='', sChar=',' → uiCount=0, uiLen=0, eOk, TRUE；
 *                         ④ sChar='' → uiCount=0, 返回 FALSE, eEmptyChar；
 *                         ⑤ sIn=';;;', sChar=';' → uiCount=3。
 *==============================================================================*)

(*-----------------------------------------------------------------------------
 * 枚举: E_DL_StrCountErr（字符计数错误码，归属 DL_Base，与本件同文件，全库唯一属主）
 *----------------------------------------------------------------------------*)
TYPE E_DL_StrCountErr :
(
    eOk        := 0,   // 信息级：统计完成 / Info: counting completed
    eEmptyChar := 1    // 故障级：目标字符为空串，统计无意义 / Fault: target character empty, counting meaningless
);
END_TYPE

FUNCTION FC_DL_StringCountChar : BOOL
VAR_INPUT
    sIn   : STRING(255);   // 被扫描字符串 [-] / Scanned string
    sChar : STRING(255);   // 目标字符源（取首字符） [-] / Target character source, first char taken
END_VAR
VAR_OUTPUT
    uiCount : UINT;        // 出现次数 [次] / Occurrence count [times]
    uiLen   : UINT;        // 扫描字符数 [字符] / Scanned character count [chars]
    eErrCode: E_DL_StrCountErr; // 错误码出口 [-] / Error code outlet
END_VAR
VAR
    _sOne   : STRING(255); // 归一后的单字符串 [-] / Normalized single character string
    _sCur   : STRING(255); // 当前扫描到的单字符 [-] / Current single character under scan
    _udLen  : UDINT;       // 输入字符数（LEN 原生宽度） [字符] / Input length in native width [chars]
    _udI    : UDINT;       // 扫描位置（1 基） [-] / Scan position, 1-based
    _uiHit  : UINT;        // 命中累加器 [次] / Hit accumulator [times]
END_VAR
VAR CONSTANT
    DL_SCC_LEN_MAX : UINT := 255;    // 缓冲上限（STRING(255) 契约） [字符] / Buffer ceiling [chars]
    DL_SCC_START   : UDINT := 1;     // 字符串起始位置（IEC 1 基） [-] / String start position, 1-based
    DL_SCC_ONE_LEN : UDINT := 1;     // 单字符长度常量 [字符] / Single character length constant [chars]
    DL_SCC_HIT_ONE : UDINT := 1;     // FIND 命中首位的比较值 [-] / Compare value for first-position hit
END_VAR

(* —— 段 0：出口预置安全值 —— *)
FC_DL_StringCountChar := FALSE;                    // 返回值预置无效 / Return preset invalid
uiCount   := 0;                                    // 计数哨兵 0 / Count sentinel
uiLen     := 0;                                    // 长度哨兵 0 / Length sentinel
eErrCode  := E_DL_StrCountErr.eEmptyChar;          // 预置最严码 / Preset strictest code

(* —— 段 1：目标字符域闸（空串无统计意义） —— *)
IF LEN(sChar) = 0 THEN
    RETURN;                                        // 保持故障码与哨兵 / Keep fault code and sentinel
END_IF

(* —— 段 2：归一为目标单字符 —— *)
_sOne := LEFT(sChar, DL_SCC_ONE_LEN);               // 取首字符（1 基索引） / Take first character, 1-based

(* —— 段 3：实测长度并钳位（缓冲可表性反算） —— *)
_udLen := LEN(sIn);                                // 输入字符数 / Input length
IF _udLen > UINT_TO_UDINT(DL_SCC_LEN_MAX) THEN
    _udLen := UINT_TO_UDINT(DL_SCC_LEN_MAX);       // 超上限钳位，保证扫描有界 / Clamp to keep scan bounded
END_IF
uiLen := UDINT_TO_UINT(_udLen);                    // 输出扫描字符数 / Export scanned length

(* —— 段 4：空串早退（零命中，仍是成功结果） —— *)
IF _udLen = 0 THEN
    eErrCode := E_DL_StrCountErr.eOk;              // 信息级成功（零命中） / Info success, zero hits
    FC_DL_StringCountChar := TRUE;
    RETURN;
END_IF

(* —— 段 5：逐字符扫描（单字符等值判定：FIND(单字符, 实测) = 1） —— *)
_uiHit := 0;                                       // 累加器清零 / Clear accumulator
_udI   := DL_SCC_START;                            // 起算位置 1 / Start at position one
WHILE _udI <= _udLen DO
    _sCur := MID(sIn, DL_SCC_ONE_LEN, _udI);       // 取第 i 个字符（1 基） / Take i-th character, 1-based
    IF FIND(_sOne, _sCur) = DL_SCC_HIT_ONE THEN
        _uiHit := _uiHit + 1;                      // 命中累加 / Accumulate one hit
    END_IF
    _udI := _udI + 1;                              // 位置步进 / Advance position
END_WHILE

(* —— 段 6：结果复检（命中数不得超过扫描长度） —— *)
IF _uiHit > uiLen THEN
    uiCount  := 0;                                 // 复检失败回哨兵 / Recheck failed: sentinel
    eErrCode := E_DL_StrCountErr.eEmptyChar;       // 保持故障级（内部不一致不入正常出口） / Keep fault-level
    RETURN;
END_IF

uiCount  := _uiHit;                                // 导出命中数 / Export hit count
eErrCode := E_DL_StrCountErr.eOk;                  // 信息级成功 / Info success
FC_DL_StringCountChar := TRUE;                     // 统计可信 / Counting trustworthy

END_FUNCTION

(* ---- FC_DL_StringCsvFieldEscape.st ---- *)
(*==============================================================================
 * 组件名称 (Component)  : FC_DL_StringCsvFieldEscape
 * 所属子库 (Sublibrary) : DL_Base
 * 当前版本 (Version)    : 1.0.0
 * 兼容性   (Platform)   : CODESYS 3.5+ / TwinCAT 3 / 汇川 InoProShop / 施耐德 Machine Expert
 *                         仅依赖 IEC 61131-3 标准字符串九函数（LEN / MID / CONCAT / FIND），零厂商私有库
 * 功能描述 (Function)   : CSV 单字段转义（RFC 4180 语义）。规则：
 *                           · 字段含逗号 / 双引号 / 换行时，整体用双引号包裹；
 *                           · 包裹时字段内每个双引号双写（" → ""）；
 *                           · 不含特殊字符时原样返回，不加引号（bQuoted=FALSE）。
 *                         用途：把 PLC 侧的批号 / 牌号 / 报警文本安全拼入 CSV 行。
 * 接口     (Interface)  : 输入 sIn 原始字段文本 [-]；
 *                         输出 sOut 转义结果、uiOutLen 结果字符数 [字符]、
 *                         bQuoted 是否已加引号、uiQuoteCount 字段内双引号个数 [个]、
 *                         eErrCode 错误码（E_DL_StrCsvErr）；
 *                         返回值 = bValid 转义有效标志（TRUE = sOut 可信）。
 * 边界     (Boundary)   : ① 属主边界：只转义单字段，不拼行、不加行尾 CR/LF、不转义分隔符本身。
 *                         ② 缓冲区可表性：转义后长度 = 原长 + 2（包裹引号）+ 引号数；
 *                         预估超 255 时判故障级 eBufferFull 并回哨兵空串（**绝不做静默截断**，
 *                         截断会破坏 CSV 语法，宁可报错交由调用方拆字段）。
 *                         ③ 换行检测依赖 IEC 字符串转义 $N（标准写法）。若某平台不解析该转义，
 *                         集合退化为两字符字面量，只会导致**多**加引号（CSV 语法仍合法），
 *                         不会漏引号——降级方向安全，已在本件显式声明。
 *                         ④ 空串合法：输出空串、bQuoted=FALSE、eOk。
 *                         ⑤ 零全局耦合（无 GVL / VAR_EXTERNAL / 物理地址）。
 * 分工声明 (Scope)      : 与 `FC_DL_StringSplitPair` 分工：反解析归那件、本件只做正向转义；
 *                         与 `FC_DL_StringRemoveWhitespace` 分工：空白剔除会破坏 CSV 语义，不混用。
 * 来源标签 (Source Tag) : 原创实现（无外部代码引入）
 * 码表     (Codes)      : 本件不占用全局数字码位；出口为 BOOL + STRING + 2×UINT + BOOL +
 *                         本文件内定义 enum E_DL_StrCsvErr（全库唯一）。
 * 红线自检 (Redline)    : R1 ✓ 零 GVL/VAR_EXTERNAL ｜ R2 ✓ 零 %I/%Q/%M ｜ R3 ✓ 纯 IEC 61131-3
 *                         R4 ✓ 预估长度前置校验（不静默截断）+ 扫描上界钳位 + 除零无路径 ｜ R5 ✓ 声明逐行同行双语注释
 *                         R6 N/A（纯函数无状态机） ｜ R7 N/A（无实例调用）
 * 修订历史 (Revision)   : 2026-11-23  v1.0.0  R77 首版（批次 B2 · 序号 10）
 * 验收向量 (Acceptance) : ① sIn='ABC' → sOut='ABC'（不加引号）, uiOutLen=3, bQuoted=FALSE, eOk；
 *                         ② sIn='A,B' → sOut='"A,B"'（7 字符）, uiOutLen=7, bQuoted=TRUE；
 *                         ③ sIn='A"B' → sOut='"A""B"'（7 字符）, uiQuoteCount=1, bQuoted=TRUE；
 *                         ④ sIn='' → sOut='', uiOutLen=0, bQuoted=FALSE, eOk；
 *                         ⑤ 转义后超 255 → 返回 FALSE, sOut='', eBufferFull。
 *==============================================================================*)

(*-----------------------------------------------------------------------------
 * 枚举: E_DL_StrCsvErr（CSV 字段转义错误码，归属 DL_Base，与本件同文件，全库唯一属主）
 * 分级: eBufferFull 为故障级（返回 FALSE，回哨兵空串）；其余为信息级（返回 TRUE）。
 *----------------------------------------------------------------------------*)
TYPE E_DL_StrCsvErr :
(
    eOk         := 0,   // 信息级：转义完成（含不加引号情形） / Info: escaping done, quoting included
    eQuoteAdded := 1,   // 信息级：已加引号包裹 / Info: field wrapped in quotes
    eBufferFull := 9    // 故障级：转义后超缓冲上限，拒绝静默截断 / Fault: escaped field exceeds buffer, silent truncation refused
);
END_TYPE

FUNCTION FC_DL_StringCsvFieldEscape : BOOL
VAR_INPUT
    sIn : STRING(255);   // 原始字段文本 [-] / Raw field text
END_VAR
VAR_OUTPUT
    sOut         : STRING(255); // 转义结果 [-] / Escaped result
    uiOutLen     : UINT;        // 结果字符数 [字符] / Result character count [chars]
    bQuoted      : BOOL;        // 是否已加引号 [-] / Whether the field was quoted
    uiQuoteCount : UINT;        // 字段内双引号个数 [个] / Number of double quotes inside the field
    eErrCode     : E_DL_StrCsvErr; // 错误码出口 [-] / Error code outlet
END_VAR
VAR
    _udLen    : UDINT;        // 输入字符数（钳位后） [字符] / Input length after clamping [chars]
    _udI      : UDINT;        // 扫描位置（1 基） [-] / Scan position, 1-based
    _udNeed   : UDINT;        // 转义后预估长度 [字符] / Estimated escaped length [chars]
    _uiQ      : UINT;         // 引号计数累加器 [个] / Quote counter accumulator
    _bSpecial : BOOL;         // 是否含需引号包裹的字符 [-] / Whether a character requiring quoting exists
    _sCur     : STRING(255);  // 当前单字符 [-] / Current single character
END_VAR
VAR CONSTANT
    DL_SCSV_DELIM : STRING(255) := ',';   // 字段分隔符（逗号） [-] / Field delimiter, comma
    DL_SCSV_QUOTE : STRING(255) := '"';   // 双引号字符 [-] / Double quote character
    DL_SCSV_QUOTE2: STRING(255) := '""';  // 双写引号（转义用） [-] / Doubled quote for escaping
    DL_SCSV_NL    : STRING(255) := '$N';  // 换行符（IEC 转义写法） [-] / Line feed via IEC escape
    DL_SCSV_LEN_MAX : UINT := 255;        // 缓冲上限（STRING(255) 契约） [字符] / Buffer ceiling [chars]
    DL_SCSV_START : UDINT := 1;           // 字符串起始位置（IEC 1 基） [-] / String start position, 1-based
    DL_SCSV_ONE_LEN: UDINT := 1;          // 单字符长度常量 [字符] / Single character length constant
    DL_SCSV_HIT_ONE: UDINT := 1;          // FIND 首位命中的比较值 [-] / Compare value for first-position hit
    DL_SCSV_WRAP   : UDINT := 2;          // 首尾包裹引号占位长度 [字符] / Wrapping quote pair length [chars]
END_VAR

(* —— 段 0：出口预置安全值 —— *)
FC_DL_StringCsvFieldEscape := FALSE;               // 返回值预置无效 / Return preset invalid
sOut         := '';                                // 结果哨兵空串 / Result sentinel
uiOutLen     := 0;                                 // 长度哨兵 0 / Length sentinel
bQuoted      := FALSE;                             // 加引号标志预置否 / Quote flag preset false
uiQuoteCount := 0;                                 // 引号计数哨兵 0 / Quote count sentinel
eErrCode     := E_DL_StrCsvErr.eBufferFull;        // 预置最严码 / Preset strictest code

(* —— 段 1：长度实测与上域钳位 —— *)
_udLen := LEN(sIn);                                // 输入字符数 / Input length
IF _udLen > UINT_TO_UDINT(DL_SCSV_LEN_MAX) THEN
    _udLen := UINT_TO_UDINT(DL_SCSV_LEN_MAX);      // 超上限钳位（仅为预估有界，不改变拒绝策略） / Clamp for bounded estimate
END_IF

(* —— 段 2：空串早退（合法零结果，不加引号） —— *)
IF _udLen = 0 THEN
    eErrCode := E_DL_StrCsvErr.eOk;                // 信息级成功 / Info success
    FC_DL_StringCsvFieldEscape := TRUE;            // 结果可信 / Result trustworthy
    RETURN;
END_IF

(* —— 段 3：扫描统计（是否需要包裹 + 引号个数） —— *)
_bSpecial := FALSE;                                // 特殊字符标志清零 / Clear special flag
_uiQ      := 0;                                    // 引号计数清零 / Clear quote counter
_udI      := DL_SCSV_START;
WHILE _udI <= _udLen DO
    _sCur := MID(sIn, DL_SCSV_ONE_LEN, _udI);      // 取第 i 个字符（1 基） / Take i-th character, 1-based
    IF FIND(DL_SCSV_DELIM, _sCur) > 0 THEN
        _bSpecial := TRUE;                         // 含分隔符需包裹 / Delimiter present: needs quoting
    END_IF
    IF FIND(DL_SCSV_QUOTE, _sCur) = DL_SCSV_HIT_ONE THEN
        _bSpecial := TRUE;                         // 含引号需包裹 / Quote present: needs quoting
        _uiQ      := _uiQ + 1;                     // 引号计数 / Count the quote
    END_IF
    IF FIND(DL_SCSV_NL, _sCur) > 0 THEN
        _bSpecial := TRUE;                         // 含换行需包裹 / Newline present: needs quoting
    END_IF
    _udI := _udI + 1;                              // 位置步进 / Advance position
END_WHILE

uiQuoteCount := _uiQ;                              // 导出引号个数 / Export quote count

(* —— 段 4：无需包裹 → 原样返回（早退，避免任何改写） —— *)
IF NOT _bSpecial THEN
    sOut     := sIn;                               // 原样返回 / Return as-is
    uiOutLen := UDINT_TO_UINT(LEN(sOut));          // 实测长度 / Measured length
    bQuoted  := FALSE;                             // 未加引号 / Not quoted
    eErrCode := E_DL_StrCsvErr.eOk;                // 信息级成功 / Info success
    FC_DL_StringCsvFieldEscape := TRUE;
    RETURN;
END_IF

(* —— 段 5：缓冲区可表性前置校验（预估超限即拒绝，绝不静默截断） —— *)
_udNeed := _udLen + DL_SCSV_WRAP + UINT_TO_UDINT(_uiQ);   // 原长 + 包裹 + 双写增量 / Original plus wrap plus doubling
IF _udNeed > UINT_TO_UDINT(DL_SCSV_LEN_MAX) THEN
    eErrCode := E_DL_StrCsvErr.eBufferFull;        // 故障级：缓冲不足 / Fault: buffer insufficient
    RETURN;                                        // 保持哨兵空串与返回 FALSE / Keep sentinel and FALSE
END_IF

(* —— 段 6：构造包裹串（先加首引号，逐字符双写，再加尾引号） —— *)
sOut := DL_SCSV_QUOTE;                             // 首引号 / Opening quote
_udI := DL_SCSV_START;
WHILE _udI <= _udLen DO
    _sCur := MID(sIn, DL_SCSV_ONE_LEN, _udI);      // 取第 i 个字符 / Take i-th character
    IF FIND(DL_SCSV_QUOTE, _sCur) = DL_SCSV_HIT_ONE THEN
        sOut := CONCAT(sOut, DL_SCSV_QUOTE2);      // 引号双写 / Double the quote
    ELSE
        sOut := CONCAT(sOut, _sCur);               // 普通字符直追加 / Append plain character
    END_IF
    _udI := _udI + 1;                              // 位置步进 / Advance position
END_WHILE
sOut := CONCAT(sOut, DL_SCSV_QUOTE);               // 尾引号 / Closing quote

(* —— 段 7：结果复检（长度必须等于预估，否则判缓冲不可信） —— *)
uiOutLen := UDINT_TO_UINT(LEN(sOut));              // 实测结果长度 / Measured result length
IF UDINT_TO_UINT(_udNeed) <> uiOutLen THEN
    sOut     := '';                                // 复检失败回哨兵 / Recheck failed: sentinel
    uiOutLen := 0;
    bQuoted  := FALSE;
    eErrCode := E_DL_StrCsvErr.eBufferFull;        // 故障级码 / Fault-level code
    RETURN;                                        // 返回 FALSE 保持 / Keep return FALSE
END_IF

(* —— 段 8：成功出口 —— *)
bQuoted  := TRUE;                                  // 已加引号 / Field quoted
eErrCode := E_DL_StrCsvErr.eQuoteAdded;            // 信息级：已包裹 / Info: wrapped
FC_DL_StringCsvFieldEscape := TRUE;                // 转义有效 / Escaping valid

END_FUNCTION

(* ---- FC_DL_StringIsNumeric.st ---- *)
(*==============================================================================
 * 组件名称 (Component)  : FC_DL_StringIsNumeric
 * 所属子库 (Sublibrary) : DL_Base
 * 当前版本 (Version)    : 1.0.0
 * 兼容性   (Platform)   : CODESYS 3.5+ / TwinCAT 3 / 汇川 InoProShop / 施耐德 Machine Expert
 *                         仅依赖 IEC 61131-3 标准字符串九函数（LEN / MID / FIND），零厂商私有库
 * 功能描述 (Function)   : 数值合法性校验（HMI 文本输入落盘前的语法前置闸）。
 *                         接受文法：  [sign] digits [ . digits ] [ (e|E) [sign] digits ]
 *                         逐字符扫描并用字符集常量做归类：
 *                           · 数字集 '0123456789'    → FIND(集合, 单字符) > 0
 *                           · 符号集 '+-'            → FIND(集合, 单字符) > 0
 *                           · 小数点 '.'             → FIND('.', 单字符) = 1
 *                           · 指数标记集 'eE'        → FIND(集合, 单字符) > 0
 *                         结构约束：符号仅允许出现在首位或指数标记之后；小数点至多一次
 *                         且不得出现在指数之后；指数至多一次且其前必须有尾数数字；
 *                         指数后必须至少有一位数字。任一违规判「非数值」。
 *                         本件只判语法，不做数值转换（转换归 STRING_TO_LREAL 调用方）。
 * 接口     (Interface)  : 输入 sIn 待校验字符串 [-]；
 *                         输出 bIsNumeric 是否数值 [-]、uiDigits 数字字符个数 [个]、
 *                         bHasSign 是否带符号、bHasDot 是否带小数点、bHasExp 是否带指数、
 *                         eErrCode 错误码（E_DL_StrNumErr）；
 *                         返回值 = bValid 判定可信标志（TRUE = bIsNumeric 可信）。
 * 边界     (Boundary)   : ① 属主边界：只判语法，不做取值范围 / 溢出 / NaN-Inf 字面量判定；
 *                         也不做空白的隐式剔除（调用方需先过 FC_DL_StringRemoveWhitespace）。
 *                         ② 空串判「非数值」（eEmptyInput，信息级），返回 TRUE（判定可信）。
 *                         ③ 含非法字符判「非数值」（eNotNumeric，信息级），返回 TRUE。
 *                         ④ '.5' / '5.' / '+5' / '-5' / '1e3' / '1.5E-3' 均判为数值；
 *                         'e5' / '1e' / '1e+' / '1.2.3' / '+-1' / '1e3.5' 判为非数值。
 *                         ⑤ 扫描上界取实测长度（<=255），严格有界；全索引 1 基。
 *                         ⑥ 零全局耦合（无 GVL / VAR_EXTERNAL / 物理地址）。
 * 分工声明 (Scope)      : 与 `FC_DL_StringSplitPair` / `FC_DL_StringRemoveWhitespace` 分工：
 *                         清洗与拆分归那两件，本件只判「是否数值」；数值转换归标准库。
 * 来源标签 (Source Tag) : 原创实现（无外部代码引入）
 * 码表     (Codes)      : 本件不占用全局数字码位；出口为 BOOL + 4 个 BOOL 特征位 + UINT +
 *                         本文件内定义 enum E_DL_StrNumErr（全库唯一）。
 * 红线自检 (Redline)    : R1 ✓ 零 GVL/VAR_EXTERNAL ｜ R2 ✓ 零 %I/%Q/%M ｜ R3 ✓ 纯 IEC 61131-3
 *                         R4 ✓ 字符集归类替代字符码强转 + 扫描上界钳位 + 状态互斥约束 ｜ R5 ✓ 声明逐行同行双语注释
 *                         R6 N/A（纯函数无状态机，用文法状态位） ｜ R7 N/A（无实例调用）
 * 修订历史 (Revision)   : 2026-11-23  v1.0.0  R77 首版（批次 B2 · 序号 5）
 * 验收向量 (Acceptance) : ① sIn='-12.5e3' → bIsNumeric=TRUE, uiDigits=4, bHasSign=TRUE,
 *                         bHasDot=TRUE, bHasExp=TRUE, eOk, 返回 TRUE；
 *                         ② sIn='12a3' → bIsNumeric=FALSE, eNotNumeric, 返回 TRUE；
 *                         ③ sIn='1e' → bIsNumeric=FALSE, eNotNumeric（指数后无数字）；
 *                         ④ sIn='' → bIsNumeric=FALSE, eEmptyInput, 返回 TRUE；
 *                         ⑤ sIn='007' → bIsNumeric=TRUE, uiDigits=3, eOk。
 *==============================================================================*)

(*-----------------------------------------------------------------------------
 * 枚举: E_DL_StrNumErr（数值合法性判定码，归属 DL_Base，与本件同文件，全库唯一属主）
 * 分级: 前四项为信息级（判定结果本身可信，返回 TRUE）；eInternal 为故障级。
 *----------------------------------------------------------------------------*)
TYPE E_DL_StrNumErr :
(
    eOk        := 0,   // 信息级：语法合法，判为数值 / Info: syntax legal, judged numeric
    eNotNumeric:= 1,   // 信息级：含非法字符或结构违规，判为非数值 / Info: illegal character or structure, judged non-numeric
    eEmptyInput:= 2,   // 信息级：空串，判为非数值 / Info: empty input, judged non-numeric
    eBadFormat := 3,   // 信息级：指数/尾数结构缺失 / Info: exponent or mantissa structure incomplete
    eInternal  := 9    // 故障级：内部一致性失败，判定不可信 / Fault: internal consistency failed, verdict untrustworthy
);
END_TYPE

FUNCTION FC_DL_StringIsNumeric : BOOL
VAR_INPUT
    sIn : STRING(255);   // 待校验字符串 [-] / String to validate
END_VAR
VAR_OUTPUT
    bIsNumeric : BOOL;   // 是否数值判定结果 [-] / Whether the text is numeric
    uiDigits   : UINT;   // 数字字符个数 [个] / Number of digit characters
    bHasSign   : BOOL;   // 是否出现合法符号 [-] / Whether a legal sign appeared
    bHasDot    : BOOL;   // 是否出现小数点 [-] / Whether a decimal point appeared
    bHasExp    : BOOL;   // 是否出现指数标记 [-] / Whether an exponent mark appeared
    eErrCode   : E_DL_StrNumErr; // 错误码出口 [-] / Error code outlet
END_VAR
VAR
    _udLen          : UDINT;      // 输入字符数（钳位后） [字符] / Input length after clamping [chars]
    _udI            : UDINT;      // 扫描位置（1 基） [-] / Scan position, 1-based
    _sCur           : STRING(255);// 当前单字符 [-] / Current single character
    _bSeenMantDigit : BOOL;       // 尾数已见数字 [-] / Mantissa digit seen
    _bSeenDot       : BOOL;       // 小数点已见 [-] / Decimal point seen
    _bSeenExp       : BOOL;       // 指数标记已见 [-] / Exponent mark seen
    _bSeenExpDigit  : BOOL;       // 指数后已见数字 [-] / Digit after exponent seen
    _bAfterExp      : BOOL;       // 刚进入指数段（符号许可窗） [-] / Just entered exponent section, sign allowed window
    _bBad           : BOOL;       // 本字符违规标志 [-] / Violation flag for current character
    _uiDig          : UINT;       // 数字累加器 [个] / Digit accumulator
END_VAR
VAR CONSTANT
    DL_SIN_SET_DIGIT : STRING(255) := '0123456789';   // 数字字符集 [-] / Digit character set
    DL_SIN_SET_SIGN  : STRING(255) := '+-';           // 符号字符集 [-] / Sign character set
    DL_SIN_SET_EXP   : STRING(255) := 'eE';           // 指数标记字符集 [-] / Exponent mark character set
    DL_SIN_DOT       : STRING(255) := '.';            // 小数点字符 [-] / Decimal point character
    DL_SIN_LEN_MAX   : UINT := 255;                   // 缓冲上限（STRING(255) 契约） [字符] / Buffer ceiling [chars]
    DL_SIN_START     : UDINT := 1;                    // 字符串起始位置（IEC 1 基） [-] / String start position, 1-based
    DL_SIN_ONE_LEN   : UDINT := 1;                    // 单字符长度常量 [字符] / Single character length constant
    DL_SIN_HIT_ONE   : UDINT := 1;                    // FIND 首位命中的比较值 [-] / Compare value for first-position hit
END_VAR

(* —— 段 0：出口预置安全值 —— *)
FC_DL_StringIsNumeric := FALSE;                    // 返回值预置不可信 / Return preset untrustworthy
bIsNumeric := FALSE;                               // 判定哨兵：非数值 / Verdict sentinel: not numeric
uiDigits   := 0;                                   // 数字计数哨兵 / Digit count sentinel
bHasSign   := FALSE;                               // 符号特征预置无 / Sign feature preset false
bHasDot    := FALSE;                               // 小数点特征预置无 / Dot feature preset false
bHasExp    := FALSE;                               // 指数特征预置无 / Exponent feature preset false
eErrCode   := E_DL_StrNumErr.eInternal;            // 预置最严码 / Preset strictest code

(* —— 段 1：长度实测与上域钳位（缓冲可表性反算，扫描严格有界） —— *)
_udLen := LEN(sIn);                                // 输入字符数 / Input length
IF _udLen > UINT_TO_UDINT(DL_SIN_LEN_MAX) THEN
    _udLen := UINT_TO_UDINT(DL_SIN_LEN_MAX);       // 超上限钳位 / Clamp to ceiling
END_IF

(* —— 段 2：空串早退（判非数值，判定本身可信） —— *)
IF _udLen = 0 THEN
    eErrCode := E_DL_StrNumErr.eEmptyInput;        // 信息级：空串 / Info: empty input
    FC_DL_StringIsNumeric := TRUE;                 // 判定可信 / Verdict trustworthy
    RETURN;
END_IF

(* —— 段 3：文法状态位预清零（不含保持量，逐次判定独立） —— *)
_bSeenMantDigit := FALSE;
_bSeenDot       := FALSE;
_bSeenExp       := FALSE;
_bSeenExpDigit  := FALSE;
_bAfterExp      := FALSE;
_bBad           := FALSE;
_uiDig          := 0;
_udI            := DL_SIN_START;

(* —— 段 4：逐字符扫描与文法约束 —— *)
WHILE _udI <= _udLen DO
    _sCur := MID(sIn, DL_SIN_ONE_LEN, _udI);       // 取第 i 个字符（1 基） / Take i-th character, 1-based
    _bBad := FALSE;                                // 每字符先清违规位 / Clear violation flag per character

    IF FIND(DL_SIN_SET_DIGIT, _sCur) > 0 THEN
        (* 数字：计数，并按所处段置位尾数/指数数字位 *)
        _uiDig := _uiDig + 1;                      // 数字计数 / Digit count
        IF _bSeenExp THEN
            _bSeenExpDigit := TRUE;                // 指数段数字 / Digit inside exponent
        ELSE
            _bSeenMantDigit := TRUE;               // 尾数段数字 / Digit inside mantissa
        END_IF
        _bAfterExp := FALSE;                       // 离开符号许可窗 / Leave sign window
    ELSIF FIND(DL_SIN_SET_SIGN, _sCur) > 0 THEN
        (* 符号：仅首位或紧指数标记之后合法 *)
        IF (_udI = DL_SIN_START) OR _bAfterExp THEN
            bHasSign   := TRUE;                    // 合法符号出现 / Legal sign recorded
            _bAfterExp := FALSE;                   // 符号用掉许可窗 / Sign consumes window
        ELSE
            _bBad := TRUE;                         // 非法位置符号 / Sign in illegal position
        END_IF
    ELSIF FIND(DL_SIN_DOT, _sCur) = DL_SIN_HIT_ONE THEN
        (* 小数点：至多一次，且不得在指数之后 *)
        IF _bSeenDot OR _bSeenExp THEN
            _bBad := TRUE;                         // 重复小数点或指数后小数点 / Duplicate dot or dot after exponent
        ELSE
            _bSeenDot := TRUE;
            bHasDot   := TRUE;
            _bAfterExp := FALSE;
        END_IF
    ELSIF FIND(DL_SIN_SET_EXP, _sCur) > 0 THEN
        (* 指数标记：至多一次，其前必须有尾数数字 *)
        IF _bSeenExp OR (NOT _bSeenMantDigit) THEN
            _bBad := TRUE;                         // 重复指数或尾数缺失 / Duplicate exponent or missing mantissa
        ELSE
            _bSeenExp  := TRUE;
            bHasExp    := TRUE;
            _bAfterExp := TRUE;                    // 打开符号许可窗 / Open sign window
        END_IF
    ELSE
        _bBad := TRUE;                             // 非法字符 / Illegal character
    END_IF

    IF _bBad THEN
        bIsNumeric := FALSE;                       // 判非数值 / Judge non-numeric
        uiDigits   := _uiDig;                      // 导出已数到的位数 / Export counted digits
        eErrCode   := E_DL_StrNumErr.eNotNumeric;  // 信息级：非法字符/结构 / Info: illegal character or structure
        FC_DL_StringIsNumeric := TRUE;             // 判定可信 / Verdict trustworthy
        RETURN;                                    // 早退 / Early exit
    END_IF

    _udI := _udI + 1;                              // 位置步进 / Advance position
END_WHILE

(* —— 段 5：收尾文法校验（尾数必须有数字；指数段必须有数字） —— *)
IF NOT _bSeenMantDigit THEN
    bIsNumeric := FALSE;                           // 无尾数数字 / No mantissa digit
    uiDigits   := _uiDig;
    eErrCode   := E_DL_StrNumErr.eBadFormat;       // 信息级：结构缺失 / Info: structure incomplete
    FC_DL_StringIsNumeric := TRUE;
    RETURN;
END_IF

IF _bSeenExp AND (NOT _bSeenExpDigit) THEN
    bIsNumeric := FALSE;                           // 指数后无数字 / No digit after exponent
    uiDigits   := _uiDig;
    eErrCode   := E_DL_StrNumErr.eBadFormat;       // 信息级：结构缺失 / Info: structure incomplete
    FC_DL_StringIsNumeric := TRUE;
    RETURN;
END_IF

(* —— 段 6：成功出口（语法合法，判为数值） —— *)
bIsNumeric := TRUE;                                // 判为数值 / Judged numeric
uiDigits   := _uiDig;                              // 导出数字个数 / Export digit count
eErrCode   := E_DL_StrNumErr.eOk;                  // 信息级成功 / Info success
FC_DL_StringIsNumeric := TRUE;                     // 判定可信 / Verdict trustworthy

END_FUNCTION
